// TIA Portal project "PADRAO" (V19)

(* hardware
DEVICE "S7-1200 station_1"  S7-1200 Station
   slot 0: "Rack_0"  S7-1200 Rack  Rack  V1.0
   slot 1: "PLC_1"  CPU 1214C DC/DC/DC  6ES7 214-1AG40-0XB0  V4.4
   slot 2: "DI 8/DQ 8x24VDC_1"  6ES7 223-1BH32-0XB0  V2.0
   slot 3: "CB 1241 (RS485)"  CB 1241 (RS485)  6ES7 241-1CH30-1XB0  V1.0
   slot 3: "DI 8/DQ 8x24VDC_2"  6ES7 223-1BH32-0XB0  V2.0
DEVICE "bb02"  GSD.Device.PN
   slot 0: "Rack"  Rack  V1.0
   slot 0: "bb02"  RT  GMXa-2-Port
      slot 0: "RT"  RT
      slot 1: "bb02"  X1
         slot 1: "Port 1"  Port 1
         slot 2: "Port 2"  Port 2
   slot 1: "Status Device_1"  Status Device
      slot 0: "Status Device"  Status Device
   slot 2: "Device Control_1"  Device Control
      slot 0: "Start/Stop"  Start/Stop
      slot 1: "Reset"  Reset
   slot 3: "Mode_1"  Mode
      slot 0: "Target Mode"  Target Mode
      slot 1: "Operating Mode"  Operating Mode
   slot 4: "Flow Rate_1"  Flow Rate
      slot 0: "Nominal Flow Rate"  Nominal Flow Rate
      slot 1: "Actual Flow Rate"  Actual Flow Rate
   slot 5: "Maximal Flow Rate_1"  Maximal Flow Rate
      slot 0: "Maximal Flow Rate"  Maximal Flow Rate
   slot 9: "Metering Monitor_1"  Metering Monitor
      slot 0: "Metering Monitor"  Metering Monitor
   slot 10: "Error/Warning_1"  Error/Warning
      slot 0: "Error"  Error
      slot 1: "Warning"  Warning
   slot 11: "Strokes/Quantities_1"  Strokes/Quantities
      slot 0: "Reset Stroke Counter"  Reset Stroke Counter
      slot 1: "Reset Quantity Counter"  Reset Quantity Counter
      slot 2: "Stroke Counter"  Stroke Counter
      slot 3: "Quantity Counter"  Quantity Counter
      slot 4: "Litres Per Stroke"  Litres Per Stroke
DEVICE "bb03"  GSD.Device.PN
   slot 0: "Rack"  Rack  V1.0
   slot 0: "bb03"  RT  GMXa-2-Port
      slot 0: "RT"  RT
      slot 1: "bb03"  X1
         slot 1: "Port 1"  Port 1
         slot 2: "Port 2"  Port 2
   slot 1: "Status Device_1"  Status Device
      slot 0: "Status Device"  Status Device
   slot 2: "Device Control_1"  Device Control
      slot 0: "Start/Stop"  Start/Stop
      slot 1: "Reset"  Reset
   slot 3: "Mode_1"  Mode
      slot 0: "Target Mode"  Target Mode
      slot 1: "Operating Mode"  Operating Mode
   slot 4: "Flow Rate_1"  Flow Rate
      slot 0: "Nominal Flow Rate"  Nominal Flow Rate
      slot 1: "Actual Flow Rate"  Actual Flow Rate
   slot 5: "Maximal Flow Rate_1"  Maximal Flow Rate
      slot 0: "Maximal Flow Rate"  Maximal Flow Rate
   slot 9: "Metering Monitor_1"  Metering Monitor
      slot 0: "Metering Monitor"  Metering Monitor
   slot 10: "Error/Warning_1"  Error/Warning
      slot 0: "Error"  Error
      slot 1: "Warning"  Warning
   slot 11: "Strokes/Quantities_1"  Strokes/Quantities
      slot 0: "Reset Stroke Counter"  Reset Stroke Counter
      slot 1: "Reset Quantity Counter"  Reset Quantity Counter
      slot 2: "Stroke Counter"  Stroke Counter
      slot 3: "Quantity Counter"  Quantity Counter
      slot 4: "Litres Per Stroke"  Litres Per Stroke
DEVICE "bb04"  GSD.Device.PN
   slot 0: "Rack"  Rack  V1.0
   slot 0: "bb04"  RT  GMXa-2-Port
      slot 0: "RT"  RT
      slot 1: "bb04"  X1
         slot 1: "Port 1"  Port 1
         slot 2: "Port 2"  Port 2
   slot 1: "Status Device_1"  Status Device
      slot 0: "Status Device"  Status Device
   slot 2: "Device Control_1"  Device Control
      slot 0: "Start/Stop"  Start/Stop
      slot 1: "Reset"  Reset
   slot 3: "Mode_1"  Mode
      slot 0: "Target Mode"  Target Mode
      slot 1: "Operating Mode"  Operating Mode
   slot 4: "Flow Rate_1"  Flow Rate
      slot 0: "Nominal Flow Rate"  Nominal Flow Rate
      slot 1: "Actual Flow Rate"  Actual Flow Rate
   slot 5: "Maximal Flow Rate_1"  Maximal Flow Rate
      slot 0: "Maximal Flow Rate"  Maximal Flow Rate
   slot 9: "Metering Monitor_1"  Metering Monitor
      slot 0: "Metering Monitor"  Metering Monitor
   slot 10: "Error/Warning_1"  Error/Warning
      slot 0: "Error"  Error
      slot 1: "Warning"  Warning
   slot 11: "Strokes/Quantities_1"  Strokes/Quantities
      slot 0: "Reset Stroke Counter"  Reset Stroke Counter
      slot 1: "Reset Quantity Counter"  Reset Quantity Counter
      slot 2: "Stroke Counter"  Stroke Counter
      slot 3: "Quantity Counter"  Quantity Counter
      slot 4: "Litres Per Stroke"  Litres Per Stroke
DEVICE "bb05"  GSD.Device.PN
   slot 0: "Rack"  Rack  V1.0
   slot 0: "bb05"  RT  GMXa-2-Port
      slot 0: "RT"  RT
      slot 1: "bb05"  X1
         slot 1: "Port 1"  Port 1
         slot 2: "Port 2"  Port 2
   slot 1: "Status Device_1"  Status Device
      slot 0: "Status Device"  Status Device
   slot 2: "Device Control_1"  Device Control
      slot 0: "Start/Stop"  Start/Stop
      slot 1: "Reset"  Reset
   slot 3: "Mode_1"  Mode
      slot 0: "Target Mode"  Target Mode
      slot 1: "Operating Mode"  Operating Mode
   slot 4: "Flow Rate_1"  Flow Rate
      slot 0: "Nominal Flow Rate"  Nominal Flow Rate
      slot 1: "Actual Flow Rate"  Actual Flow Rate
   slot 5: "Maximal Flow Rate_1"  Maximal Flow Rate
      slot 0: "Maximal Flow Rate"  Maximal Flow Rate
   slot 9: "Metering Monitor_1"  Metering Monitor
      slot 0: "Metering Monitor"  Metering Monitor
   slot 10: "Error/Warning_1"  Error/Warning
      slot 0: "Error"  Error
      slot 1: "Warning"  Warning
   slot 11: "Strokes/Quantities_1"  Strokes/Quantities
      slot 0: "Reset Stroke Counter"  Reset Stroke Counter
      slot 1: "Reset Quantity Counter"  Reset Quantity Counter
      slot 2: "Stroke Counter"  Stroke Counter
      slot 3: "Quantity Counter"  Quantity Counter
      slot 4: "Litres Per Stroke"  Litres Per Stroke
DEVICE "bb01"  GSD.Device.PN
   slot 0: "Rack"  Rack  V1.0
   slot 0: "bb01"  RT  GMXa-2-Port
      slot 0: "RT"  RT
      slot 1: "bb01"  X1
         slot 1: "Port 1"  Port 1
         slot 2: "Port 2"  Port 2
   slot 1: "Status Device_1"  Status Device
      slot 0: "Status Device"  Status Device
   slot 2: "Device Control_1"  Device Control
      slot 0: "Start/Stop"  Start/Stop
      slot 1: "Reset"  Reset
   slot 3: "Mode_1"  Mode
      slot 0: "Target Mode"  Target Mode
      slot 1: "Operating Mode"  Operating Mode
   slot 4: "Flow Rate_1"  Flow Rate
      slot 0: "Nominal Flow Rate"  Nominal Flow Rate
      slot 1: "Actual Flow Rate"  Actual Flow Rate
   slot 5: "Maximal Flow Rate_1"  Maximal Flow Rate
      slot 0: "Maximal Flow Rate"  Maximal Flow Rate
   slot 9: "Metering Monitor_1"  Metering Monitor
      slot 0: "Metering Monitor"  Metering Monitor
   slot 10: "Error/Warning_1"  Error/Warning
      slot 0: "Error"  Error
      slot 1: "Warning"  Warning
   slot 11: "Strokes/Quantities_1"  Strokes/Quantities
      slot 0: "Reset Stroke Counter"  Reset Stroke Counter
      slot 1: "Reset Quantity Counter"  Reset Quantity Counter
      slot 2: "Stroke Counter"  Stroke Counter
      slot 3: "Quantity Counter"  Quantity Counter
      slot 4: "Litres Per Stroke"  Litres Per Stroke
DEVICE "bb05_1"  GSD.Device.PN
   slot 0: "Rack"  Rack  V1.0
   slot 0: "bb06"  RT  GMXa-2-Port
      slot 0: "RT"  RT
      slot 1: "bb06"  X1
         slot 1: "Port 1"  Port 1
         slot 2: "Port 2"  Port 2
   slot 1: "Status Device_1"  Status Device
      slot 0: "Status Device"  Status Device
   slot 2: "Device Control_1"  Device Control
      slot 0: "Start/Stop"  Start/Stop
      slot 1: "Reset"  Reset
   slot 3: "Mode_1"  Mode
      slot 0: "Target Mode"  Target Mode
      slot 1: "Operating Mode"  Operating Mode
   slot 4: "Flow Rate_1"  Flow Rate
      slot 0: "Nominal Flow Rate"  Nominal Flow Rate
      slot 1: "Actual Flow Rate"  Actual Flow Rate
   slot 5: "Maximal Flow Rate_1"  Maximal Flow Rate
      slot 0: "Maximal Flow Rate"  Maximal Flow Rate
   slot 9: "Metering Monitor_1"  Metering Monitor
      slot 0: "Metering Monitor"  Metering Monitor
   slot 10: "Error/Warning_1"  Error/Warning
      slot 0: "Error"  Error
      slot 1: "Warning"  Warning
   slot 11: "Strokes/Quantities_1"  Strokes/Quantities
      slot 0: "Reset Stroke Counter"  Reset Stroke Counter
      slot 1: "Reset Quantity Counter"  Reset Quantity Counter
      slot 2: "Stroke Counter"  Stroke Counter
      slot 3: "Quantity Counter"  Quantity Counter
      slot 4: "Litres Per Stroke"  Litres Per Stroke
*)

// ===== PLC "PLC_1"  CPU 1214C DC/DC/DC =====

VAR_GLOBAL   // PLC tag table "Default tag table"
   "DI_00" AT %I0.0 : Bool;
   "DI_01" AT %I0.1 : Bool;
   "DI_02" AT %I0.2 : Bool;
   "DI_03" AT %I0.3 : Bool;
   "DI_04" AT %I0.4 : Bool;
   "DI_05" AT %I0.5 : Bool;
   "DI_06" AT %I0.6 : Bool;
   "DI_07" AT %I0.7 : Bool;
   "DI_08" AT %I1.0 : Bool;
   "DI_09" AT %I1.1 : Bool;
   "DI_10" AT %I1.2 : Bool;
   "DI_11" AT %I1.3 : Bool;
   "DI_12" AT %I1.4 : Bool;
   "DI_13" AT %I1.5 : Bool;
   "DO_00" AT %Q0.0 : Bool;
   "DO_01" AT %Q0.1 : Bool;
   "DO_02" AT %Q0.2 : Bool;
   "DO_03" AT %Q0.3 : Bool;
   "DO_04" AT %Q0.4 : Bool;
   "DO_05" AT %Q0.5 : Bool;
   "DO_06" AT %Q0.6 : Bool;
   "DO_07" AT %Q0.7 : Bool;
   "DO_08" AT %Q1.0 : Bool;
   "DO_09" AT %Q1.1 : Bool;
   "System_Byte" AT %MB1 : Byte;
   "FirstScan" AT %M1.0 : Bool;
   "DiagStatusUpdate" AT %M1.1 : Bool;
   "AlwaysTRUE" AT %M1.2 : Bool;
   "AlwaysFALSE" AT %M1.3 : Bool;
   "Clock_Byte" AT %MB0 : Byte;
   "Clock_10Hz" AT %M0.0 : Bool;
   "Clock_5Hz" AT %M0.1 : Bool;
   "Clock_2.5Hz" AT %M0.2 : Bool;
   "Clock_2Hz" AT %M0.3 : Bool;
   "Clock_1.25Hz" AT %M0.4 : Bool;
   "Clock_1Hz" AT %M0.5 : Bool;
   "Clock_0.625Hz" AT %M0.6 : Bool;
   "Clock_0.5Hz" AT %M0.7 : Bool;
   "EmergenciaAcionada" AT %M2.0 : Bool;
   "FaltaFase" AT %M2.1 : Bool;
   "SinalTriturador1" AT %M2.2 : Bool;
   "SinalTriturador2" AT %M2.3 : Bool;
   "SinalMisturador1" AT %M2.4 : Bool;
   "SinalMisturador2" AT %M2.5 : Bool;
   "PulsoMedidor1" AT %M3.3 : Bool;
   "PulsoMedidor2" AT %M3.4 : Bool;
   "PulsoMedidor3" AT %M3.5 : Bool;
   "SistemaHabilitado" AT %M3.6 : Bool;
   "Sirene" AT %M3.7 : Bool;
   "FatorCorrecaoTanque1" AT %MD108 : Real;
   "AI_01" AT %IW64 : Word;
   "AI_02" AT %IW66 : Word;
   "ResetGeral" AT %M4.0 : Bool;
   "VolumePulso1" AT %MD160 : Real;
   "VolumePulso2" AT %MD164 : Real;
   "VolumePulso3" AT %MD172 : Real;
   "NivelBaixoTQ1" AT %M4.1 : Bool;
   "SP_NivelMinimoTanque1" AT %MD184 : Real;
   "StatusFalha" AT %MW192 : Int;
   "FalhaBomba01" AT %M4.5 : Bool;
   "FalhaBomba02" AT %M4.6 : Bool;
   "FalhaBomba03" AT %M4.7 : Bool;
   "FalhaBomba04" AT %M5.0 : Bool;
   "FalhaBomba05" AT %M5.1 : Bool;
   "FatorCorrecaoTanque2" AT %MD112 : Real;
   "SP_NivelMinimoTanque2" AT %MD152 : Real;
   "NivelBaixoTQ2" AT %M7.5 : Bool;
   "LigaValv04" AT %M7.6 : Bool;
   "LigaValv05" AT %M7.7 : Bool;
   "VolumePulso4" AT %MD100 : Real;
   "SP_Dosagem1" AT %MD168 : Real;
   "SP_Dosagem2" AT %MD176 : Real;
   "SP_Dosagem3" AT %MD180 : Real;
   "SP_Dosagem4" AT %MD188 : Real;
   "SP_Dosagem5" AT %MD194 : Real;
   "PulsoMedidor4" AT %M8.2 : Bool;
   "PulsoMedidor5" AT %M8.3 : Bool;
   "FaltaFluxo01" AT %M2.6 : Bool;
   "FaltaFluxo02" AT %M2.7 : Bool;
   "FaltaFluxo03" AT %M3.0 : Bool;
   "FaltaFluxo04" AT %M3.1 : Bool;
   "FaltaFluxo05" AT %M3.2 : Bool;
   "VolumePulso5" AT %MD104 : Real;
   "LigaValv03" AT %M8.0 : Bool;
   "LigaValv06" AT %M8.1 : Bool;
   "RetValvAberta3" AT %M8.5 : Bool;
   "RetValvAberta4" AT %M8.6 : Bool;
   "RetValvAberta5" AT %M8.7 : Bool;
   "RetValvAberta6" AT %M9.0 : Bool;
   "FalhaRetornoValvAberta3" AT %M9.1 : Bool;
   "FalhaRetornoValvAberta4" AT %M9.2 : Bool;
   "FalhaRetornoValvAberta5" AT %M9.3 : Bool;
   "BombaMax1" AT %M4.2 : Bool;
   "BombaMax2" AT %M4.3 : Bool;
   "BombaMax3" AT %M4.4 : Bool;
   "BombaMax4" AT %M5.3 : Bool;
   "BombaMax5" AT %M5.4 : Bool;
   "MedidorEstragado1" AT %M5.5 : Bool;
   "MedidorEstragado2" AT %M5.6 : Bool;
   "MedidorEstragado3" AT %M5.7 : Bool;
   "MedidorEstragado4" AT %M6.0 : Bool;
   "MedidorEstragado5" AT %M6.1 : Bool;
   "IniciaCalibracao1" AT %M6.3 : Bool;
   "IniciaCalibracao2" AT %M6.4 : Bool;
   "IniciaCalibracao3" AT %M6.5 : Bool;
   "IniciaCalibracao4" AT %M6.6 : Bool;
   "IniciaCalibracao5" AT %M6.7 : Bool;
   "BombaMax6" AT %M7.1 : Bool;
   "FalhaBomba06" AT %M5.2 : Bool;
   "FalhaRetornoValvAberta6" AT %M9.4 : Bool;
   "FaltaFluxo06" AT %M6.2 : Bool;
   "VolumePulso6" AT %MD116 : Real;
   "IniciaCalibracao6" AT %M7.0 : Bool;
   "MedidorEstragado6" AT %M7.2 : Bool;
   "PulsoMedidor6" AT %M8.4 : Bool;
   "SP_Dosagem6" AT %MD198 : Real;
   "SP_NivelMuitoBaixoTanque1" AT %MD120 : Real;
   "SP_NivelMuitoBaixoTanque2" AT %MD124 : Real;
   "NivelMuitoBaixoTQ1" AT %M7.3 : Bool;
   "NivelMuitoBaixoTQ2" AT %M7.4 : Bool;
   "OffSetTQ1" AT %MD128 : Real;
   "OffSetTQ2" AT %MD132 : Real;
   "CircunferenciaTQ1" AT %MD136 : Real;
   "CircunferenciaTQ2" AT %MD140 : Real;
   "StatusBombaEspelho" AT %MD144 : DInt;
   "DataEspelho" AT %MD148 : DInt;
   "HoraEspelho" AT %MD156 : DInt;
   "DI_14" AT %I8.0 : Bool;
   "DI_15" AT %I8.1 : Bool;
   "DI_16" AT %I8.2 : Bool;
   "DI_17" AT %I8.3 : Bool;
   "DI_18" AT %I8.4 : Bool;
   "DI_19" AT %I8.5 : Bool;
   "DI_20" AT %I8.6 : Bool;
   "DI_21" AT %I8.7 : Bool;
   "SP_DelayFinal1" AT %MD202 : Time;
   "SP_DelayFinal2" AT %MD206 : Time;
   "SP_DelayFinal3" AT %MD210 : Time;
   "SP_DelayFinal4" AT %MD214 : Time;
   "SP_DelayFinal5" AT %MD218 : Time;
   "SP_DelayFinal6" AT %MD222 : Time;
   "FalhaRetBomba1" AT %M9.5 : Bool;
   "FalhaRetBomba2" AT %M9.6 : Bool;
   "FalhaRetBomba3" AT %M9.7 : Bool;
   "FalhaRetBomba4" AT %M10.0 : Bool;
   "FalhaRetBomba5" AT %M10.1 : Bool;
   "FalhaRetBomba6" AT %M10.2 : Bool;
   "QuedaEnergia" AT %M10.3 : Bool;
   "Frequencia1" AT %MD246 : Real;
   "SP_DelayIniciaPID" AT %MD242 : Time;
   "Frequencia2" AT %MD250 : Real;
   "Frequencia3" AT %MD254 : Real;
   "Frequencia4" AT %MD258 : Real;
   "Frequencia5" AT %MD262 : Real;
   "Frequencia6" AT %MD300 : Real;
   "SP_DelayColaFreq" AT %MD12 : Time;
END_VAR

// folder: Common

TYPE "typeDiagnostics"
TITLE = typeDiagnostics
// Provides a structure for detailed diagnostics
   STRUCT
      status : Word;   // Status of the block or error identification when error occurred
      subfunctionStatus : DWord;   // Status or return value of called FBs, FCs and system blocks
      stateNumber : DInt;   // State in the state machine of the block where the error occurred
   END_STRUCT;
END_TYPE

// folder: LMQTT

TYPE "LMQTT_typeConnParam"
TITLE = LMQTT_typeConnParams
// Specifies connection parameters for the mqtt connection
   STRUCT
      hwId : Hw_Any;   // Hardware identifier of the interface. 0: interface is selected automatically
      connId : Conn_Ouc := 1;   // Unique connection identifier (1..4095)
      broker : String;   // Hostname or IP address of broker
      port : UInt := 1883;   // Port on the broker
      tls : Struct   // Parameters for TLS encryption
         enableTls : Bool;   // TRUE: Enables TLS, FALSE: disable TLS
         validateServerIdentity : Bool;   // TRUE: Validate server certificate, FALSE: No validation of server certificate
         brokerCert : UDInt;   // ID of the broker's certificate in TIA Portal
         clientCert : UDInt;   // ID of the client's certificate in TIA Portal
      END_STRUCT;
      keepAlive : UInt;   // Keepalive mechanism for MQTT in seconds. 0: disabled.
   END_STRUCT;
END_TYPE

// folder: DB

DATA_BLOCK "RelatorioUnificado"   // DB1
{ S7_Optimized_Access := 'TRUE' }
VERSION : 0.1
   VAR RETAIN
      Diario : Array[1..20] of Real;
      Totalizador : Array[1..20] of Real;
      DosagemAtual : Array[1..20] of Real;
   END_VAR
BEGIN
END_DATA_BLOCK

DATA_BLOCK "InputClp_DB"   // DB2
{ S7_Optimized_Access := 'TRUE' }
VERSION : 0.1
// stored: InstanceOfName InputClp
"InputClp"
BEGIN
END_DATA_BLOCK

DATA_BLOCK "NivelTanque1"   // DB3
{ S7_Optimized_Access := 'TRUE' }
VERSION : 0.1
// stored: InstanceOfName NivelTanque
"NivelTanque"
BEGIN
END_DATA_BLOCK

DATA_BLOCK "InputClp_DB2"   // DB4
{ S7_Optimized_Access := 'TRUE' }
VERSION : 0.1
// stored: InstanceOfName InputClp
"InputClp"
BEGIN
END_DATA_BLOCK

DATA_BLOCK "OutputClp_DB"   // DB5
{ S7_Optimized_Access := 'TRUE' }
VERSION : 0.1
// stored: InstanceOfName OutputClp
"OutputClp"
BEGIN
END_DATA_BLOCK

DATA_BLOCK "NivelTanque2"   // DB6
{ S7_Optimized_Access := 'TRUE' }
VERSION : 0.1
// stored: InstanceOfName NivelTanque
"NivelTanque"
BEGIN
END_DATA_BLOCK

DATA_BLOCK "DosagemContinua_DB1"   // DB7
{ S7_Optimized_Access := 'TRUE' }
VERSION : 0.1
// stored: InstanceOfName DosagemContinua
"DosagemContinua"
BEGIN
END_DATA_BLOCK

DATA_BLOCK "RegistradorMedidor_DB1"   // DB8
{ S7_Optimized_Access := 'TRUE' }
VERSION : 0.1
// stored: InstanceOfName RegistradorMedidor
"RegistradorMedidor"
BEGIN
END_DATA_BLOCK

DATA_BLOCK "DosagemContinua_DB2"   // DB9
{ S7_Optimized_Access := 'TRUE' }
VERSION : 0.1
// stored: InstanceOfName DosagemContinua
"DosagemContinua"
BEGIN
END_DATA_BLOCK

DATA_BLOCK "RegistradorMedidor_DB2"   // DB10
{ S7_Optimized_Access := 'TRUE' }
VERSION : 0.1
// stored: InstanceOfName RegistradorMedidor
"RegistradorMedidor"
BEGIN
END_DATA_BLOCK

DATA_BLOCK "DosagemContinua_DB3"   // DB11
{ S7_Optimized_Access := 'TRUE' }
VERSION : 0.1
// stored: InstanceOfName DosagemContinua
"DosagemContinua"
BEGIN
END_DATA_BLOCK

DATA_BLOCK "RegistradorMedidor_DB3"   // DB12
{ S7_Optimized_Access := 'TRUE' }
VERSION : 0.1
// stored: InstanceOfName RegistradorMedidor
"RegistradorMedidor"
BEGIN
END_DATA_BLOCK

DATA_BLOCK "DosagemContinua_DB4"   // DB13
{ S7_Optimized_Access := 'TRUE' }
VERSION : 0.1
// stored: InstanceOfName DosagemContinua
"DosagemContinua"
BEGIN
END_DATA_BLOCK

DATA_BLOCK "RelatorioSAPI"   // DB14
{ S7_Optimized_Access := 'TRUE' }
VERSION : 0.1
   VAR RETAIN
      Hora : Array[1..200] of Real;
      TotalTempoBomba : Array[1..20] of DInt;
      TotalTempoSinal : Array[1..20] of DInt;
      TotalAcionamentosSinal : Array[1..20] of DInt;
      TotalAcionamentosBBA : Array[1..20] of DInt;
      auxPulsoClock : Array[1..40] of Bool;
      auxNegaSinal : Array[1..20] of Bool;
      auxNegaBomba : Array[1..20] of Bool;
      StatusINT : Int := -1;
      StatusReal : Real := -1.0;
   END_VAR
   VAR
      GravaFTP : Bool;
      EnviaFTP : Bool;
      TesteGrava : Bool;
      TesteEnvia : Bool;
      TesteSet : Bool;
   END_VAR
BEGIN
   Hora[1] := -1.0;
   Hora[2] := -1.0;
   Hora[3] := -1.0;
   Hora[4] := -1.0;
   Hora[5] := -1.0;
   Hora[6] := -1.0;
   Hora[7] := -1.0;
   Hora[8] := -1.0;
   Hora[9] := -1.0;
   Hora[10] := -1.0;
   Hora[11] := -1.0;
   Hora[12] := -1.0;
   Hora[13] := -1.0;
   Hora[14] := -1.0;
   Hora[15] := -1.0;
   Hora[16] := -1.0;
   Hora[17] := -1.0;
   Hora[18] := -1.0;
   Hora[19] := -1.0;
   Hora[20] := -1.0;
   Hora[21] := -1.0;
   Hora[22] := -1.0;
   Hora[23] := -1.0;
   Hora[24] := -1.0;
   Hora[25] := -1.0;
   Hora[26] := -1.0;
   Hora[27] := -1.0;
   Hora[28] := -1.0;
   Hora[29] := -1.0;
   Hora[30] := -1.0;
   Hora[31] := -1.0;
   Hora[32] := -1.0;
   Hora[33] := -1.0;
   Hora[34] := -1.0;
   Hora[35] := -1.0;
   Hora[36] := -1.0;
   Hora[37] := -1.0;
   Hora[38] := -1.0;
   Hora[39] := -1.0;
   Hora[40] := -1.0;
   Hora[41] := -1.0;
   Hora[42] := -1.0;
   Hora[43] := -1.0;
   Hora[44] := -1.0;
   Hora[45] := -1.0;
   Hora[46] := -1.0;
   Hora[47] := -1.0;
   Hora[48] := -1.0;
   Hora[49] := -1.0;
   Hora[50] := -1.0;
   Hora[51] := -1.0;
   Hora[52] := -1.0;
   Hora[53] := -1.0;
   Hora[54] := -1.0;
   Hora[55] := -1.0;
   Hora[56] := -1.0;
   Hora[57] := -1.0;
   Hora[58] := -1.0;
   Hora[59] := -1.0;
   Hora[60] := -1.0;
   Hora[61] := -1.0;
   Hora[62] := -1.0;
   Hora[63] := -1.0;
   Hora[64] := -1.0;
   Hora[65] := -1.0;
   Hora[66] := -1.0;
   Hora[67] := -1.0;
   Hora[68] := -1.0;
   Hora[69] := -1.0;
   Hora[70] := -1.0;
   Hora[71] := -1.0;
   Hora[72] := -1.0;
   Hora[73] := -1.0;
   Hora[74] := -1.0;
   Hora[75] := -1.0;
   Hora[76] := -1.0;
   Hora[77] := -1.0;
   Hora[78] := -1.0;
   Hora[79] := -1.0;
   Hora[80] := -1.0;
   Hora[81] := -1.0;
   Hora[82] := -1.0;
   Hora[83] := -1.0;
   Hora[84] := -1.0;
   Hora[85] := -1.0;
   Hora[86] := -1.0;
   Hora[87] := -1.0;
   Hora[88] := -1.0;
   Hora[89] := -1.0;
   Hora[90] := -1.0;
   Hora[91] := -1.0;
   Hora[92] := -1.0;
   Hora[93] := -1.0;
   Hora[94] := -1.0;
   Hora[95] := -1.0;
   Hora[96] := -1.0;
   Hora[97] := -1.0;
   Hora[98] := -1.0;
   Hora[99] := -1.0;
   Hora[100] := -1.0;
   Hora[101] := -1.0;
   Hora[102] := -1.0;
   Hora[103] := -1.0;
   Hora[104] := -1.0;
   Hora[105] := -1.0;
   Hora[106] := -1.0;
   Hora[107] := -1.0;
   Hora[108] := -1.0;
   Hora[109] := -1.0;
   Hora[110] := -1.0;
   Hora[111] := -1.0;
   Hora[112] := -1.0;
   Hora[113] := -1.0;
   Hora[114] := -1.0;
   Hora[115] := -1.0;
   Hora[116] := -1.0;
   Hora[117] := -1.0;
   Hora[118] := -1.0;
   Hora[119] := -1.0;
   Hora[120] := -1.0;
   Hora[121] := -1.0;
   Hora[122] := -1.0;
   Hora[123] := -1.0;
   Hora[124] := -1.0;
   Hora[125] := -1.0;
   Hora[126] := -1.0;
   Hora[127] := -1.0;
   Hora[128] := -1.0;
   Hora[129] := -1.0;
   Hora[130] := -1.0;
   Hora[131] := -1.0;
   Hora[132] := -1.0;
   Hora[133] := -1.0;
   Hora[134] := -1.0;
   Hora[135] := -1.0;
   Hora[136] := -1.0;
   Hora[137] := -1.0;
   Hora[138] := -1.0;
   Hora[139] := -1.0;
   Hora[140] := -1.0;
   Hora[141] := -1.0;
   Hora[142] := -1.0;
   Hora[143] := -1.0;
   Hora[144] := -1.0;
   Hora[145] := -1.0;
   Hora[146] := -1.0;
   Hora[147] := -1.0;
   Hora[148] := -1.0;
   Hora[149] := -1.0;
   Hora[150] := -1.0;
   Hora[151] := -1.0;
   Hora[152] := -1.0;
   Hora[153] := -1.0;
   Hora[154] := -1.0;
   Hora[155] := -1.0;
   Hora[156] := -1.0;
   Hora[157] := -1.0;
   Hora[158] := -1.0;
   Hora[159] := -1.0;
   Hora[160] := -1.0;
   Hora[161] := -1.0;
   Hora[162] := -1.0;
   Hora[163] := -1.0;
   Hora[164] := -1.0;
   Hora[165] := -1.0;
   Hora[166] := -1.0;
   Hora[167] := -1.0;
   Hora[168] := -1.0;
   Hora[169] := -1.0;
   Hora[170] := -1.0;
   Hora[171] := -1.0;
   Hora[172] := -1.0;
   Hora[173] := -1.0;
   Hora[174] := -1.0;
   Hora[175] := -1.0;
   Hora[176] := -1.0;
   Hora[177] := -1.0;
   Hora[178] := -1.0;
   Hora[179] := -1.0;
   Hora[180] := -1.0;
   Hora[181] := -1.0;
   Hora[182] := -1.0;
   Hora[183] := -1.0;
   Hora[184] := -1.0;
   Hora[185] := -1.0;
   Hora[186] := -1.0;
   Hora[187] := -1.0;
   Hora[188] := -1.0;
   Hora[189] := -1.0;
   Hora[190] := -1.0;
   Hora[191] := -1.0;
   Hora[192] := -1.0;
   Hora[193] := -1.0;
   Hora[194] := -1.0;
   Hora[195] := -1.0;
   Hora[196] := -1.0;
   Hora[197] := -1.0;
   Hora[198] := -1.0;
   Hora[199] := -1.0;
   Hora[200] := -1.0;
END_DATA_BLOCK

DATA_BLOCK "RegistradorMedidor_DB4"   // DB15
{ S7_Optimized_Access := 'TRUE' }
VERSION : 0.1
// stored: InstanceOfName RegistradorMedidor
"RegistradorMedidor"
BEGIN
END_DATA_BLOCK

DATA_BLOCK "InterfaceProfi1"   // DB16
{ S7_Optimized_Access := 'TRUE' }
AUTHOR : kellerc
FAMILY : GammaX
NAME : Basic
VERSION : 1.0
// stored: InstanceOfName FBGammaX_1200
"FBGammaX_1200"
BEGIN
END_DATA_BLOCK

DATA_BLOCK "DosagemContinua_DB5"   // DB17
{ S7_Optimized_Access := 'TRUE' }
VERSION : 0.1
// stored: InstanceOfName DosagemContinua
"DosagemContinua"
BEGIN
END_DATA_BLOCK

DATA_BLOCK "InterfaceProfi2"   // DB18
{ S7_Optimized_Access := 'TRUE' }
AUTHOR : kellerc
FAMILY : GammaX
NAME : Basic
VERSION : 1.0
// stored: InstanceOfName FBGammaX_1200
"FBGammaX_1200"
BEGIN
END_DATA_BLOCK

DATA_BLOCK "InterfaceProfi3"   // DB19
{ S7_Optimized_Access := 'TRUE' }
AUTHOR : kellerc
FAMILY : GammaX
NAME : Basic
VERSION : 1.0
// stored: InstanceOfName FBGammaX_1200
"FBGammaX_1200"
BEGIN
END_DATA_BLOCK

DATA_BLOCK "InterfaceProfi4"   // DB20
{ S7_Optimized_Access := 'TRUE' }
AUTHOR : kellerc
FAMILY : GammaX
NAME : Basic
VERSION : 1.0
// stored: InstanceOfName FBGammaX_1200
"FBGammaX_1200"
BEGIN
END_DATA_BLOCK

DATA_BLOCK "InterfaceProfi5"   // DB21
{ S7_Optimized_Access := 'TRUE' }
AUTHOR : kellerc
FAMILY : GammaX
NAME : Basic
VERSION : 1.0
// stored: InstanceOfName FBGammaX_1200
"FBGammaX_1200"
BEGIN
END_DATA_BLOCK

DATA_BLOCK "RegistradorMedidor_DB5"   // DB22
{ S7_Optimized_Access := 'TRUE' }
VERSION : 0.1
// stored: InstanceOfName RegistradorMedidor
"RegistradorMedidor"
BEGIN
END_DATA_BLOCK

DATA_BLOCK "DosagemContinua_DB6"   // DB23
{ S7_Optimized_Access := 'TRUE' }
VERSION : 0.1
// stored: InstanceOfName DosagemContinua
"DosagemContinua"
BEGIN
END_DATA_BLOCK

DATA_BLOCK "RegistradorMedidor_DB6"   // DB24
{ S7_Optimized_Access := 'TRUE' }
VERSION : 0.1
// stored: InstanceOfName RegistradorMedidor
"RegistradorMedidor"
BEGIN
END_DATA_BLOCK

DATA_BLOCK "InterfaceProfi6"   // DB31
{ S7_Optimized_Access := 'TRUE' }
AUTHOR : kellerc
FAMILY : GammaX
NAME : Basic
VERSION : 1.0
// stored: InstanceOfName FBGammaX_1200
"FBGammaX_1200"
BEGIN
END_DATA_BLOCK

DATA_BLOCK "DataTime"   // DB48
{ S7_Optimized_Access := 'TRUE' }
VERSION : 0.1
   VAR RETAIN
      DataHora : DTL;
      IHM : Array[0..6] of Word;
   END_VAR
BEGIN
END_DATA_BLOCK

DATA_BLOCK "SetDbSapi_DB"   // DB87
{ S7_Optimized_Access := 'TRUE' }
VERSION : 0.1
// stored: InstanceOfName SetDbSapi
"SetDbSapi"
BEGIN
END_DATA_BLOCK

// folder: System blocks/Program resources

DATA_BLOCK "TON_FalhaRetornoValv3"   // DB25
{ S7_Optimized_Access := 'TRUE' }
AUTHOR : Simatic
FAMILY : IEC
NAME : IEC_TMR
VERSION : 1.0
// stored: InstanceOfName IEC_TIMER
"IEC_TIMER"
BEGIN
END_DATA_BLOCK

DATA_BLOCK "TON_FalhaRetornoValv4"   // DB26
{ S7_Optimized_Access := 'TRUE' }
AUTHOR : Simatic
FAMILY : IEC
NAME : IEC_TMR
VERSION : 1.0
// stored: InstanceOfName IEC_TIMER
"IEC_TIMER"
BEGIN
END_DATA_BLOCK

DATA_BLOCK "TON_FalhaRetornoValv5"   // DB27
{ S7_Optimized_Access := 'TRUE' }
AUTHOR : Simatic
FAMILY : IEC
NAME : IEC_TMR
VERSION : 1.0
// stored: InstanceOfName IEC_TIMER
"IEC_TIMER"
BEGIN
END_DATA_BLOCK

DATA_BLOCK "TON_FalhaRetornoValv6"   // DB28
{ S7_Optimized_Access := 'TRUE' }
AUTHOR : Simatic
FAMILY : IEC
NAME : IEC_TMR
VERSION : 1.0
// stored: InstanceOfName IEC_TIMER
"IEC_TIMER"
BEGIN
END_DATA_BLOCK

DATA_BLOCK "TON_DelayIniciaPID1"   // DB29
{ S7_Optimized_Access := 'TRUE' }
AUTHOR : Simatic
FAMILY : IEC
NAME : IEC_TMR
VERSION : 1.0
// stored: InstanceOfName IEC_TIMER
"IEC_TIMER"
BEGIN
END_DATA_BLOCK

DATA_BLOCK "TON_DelayIniciaPID2"   // DB30
{ S7_Optimized_Access := 'TRUE' }
AUTHOR : Simatic
FAMILY : IEC
NAME : IEC_TMR
VERSION : 1.0
// stored: InstanceOfName IEC_TIMER
"IEC_TIMER"
BEGIN
END_DATA_BLOCK

DATA_BLOCK "TON_DelayIniciaPID3"   // DB32
{ S7_Optimized_Access := 'TRUE' }
AUTHOR : Simatic
FAMILY : IEC
NAME : IEC_TMR
VERSION : 1.0
// stored: InstanceOfName IEC_TIMER
"IEC_TIMER"
BEGIN
END_DATA_BLOCK

DATA_BLOCK "TON_DelayIniciaPID4"   // DB33
{ S7_Optimized_Access := 'TRUE' }
AUTHOR : Simatic
FAMILY : IEC
NAME : IEC_TMR
VERSION : 1.0
// stored: InstanceOfName IEC_TIMER
"IEC_TIMER"
BEGIN
END_DATA_BLOCK

DATA_BLOCK "TON_DelayIniciaPID5"   // DB34
{ S7_Optimized_Access := 'TRUE' }
AUTHOR : Simatic
FAMILY : IEC
NAME : IEC_TMR
VERSION : 1.0
// stored: InstanceOfName IEC_TIMER
"IEC_TIMER"
BEGIN
END_DATA_BLOCK

DATA_BLOCK "TON_DelayIniciaPID6"   // DB35
{ S7_Optimized_Access := 'TRUE' }
AUTHOR : Simatic
FAMILY : IEC
NAME : IEC_TMR
VERSION : 1.0
// stored: InstanceOfName IEC_TIMER
"IEC_TIMER"
BEGIN
END_DATA_BLOCK

DATA_BLOCK "TON_ResetQuedaEnergia"   // DB42
{ S7_Optimized_Access := 'TRUE' }
AUTHOR : Simatic
FAMILY : IEC
NAME : IEC_TMR
VERSION : 1.0
// stored: InstanceOfName IEC_TIMER
"IEC_TIMER"
BEGIN
END_DATA_BLOCK

DATA_BLOCK "TOF_ResetGeral"   // DB43
{ S7_Optimized_Access := 'TRUE' }
AUTHOR : Simatic
FAMILY : IEC
NAME : IEC_TMR
VERSION : 1.0
// stored: InstanceOfName IEC_TIMER
"IEC_TIMER"
BEGIN
END_DATA_BLOCK

DATA_BLOCK "ModbusTimer1"   // DB46
{ S7_Optimized_Access := 'TRUE' }
AUTHOR : Simatic
FAMILY : IEC
NAME : IEC_TMR
VERSION : 1.0
// stored: InstanceOfName IEC_TIMER
"IEC_TIMER"
BEGIN
END_DATA_BLOCK

DATA_BLOCK "ContadorFalha1"   // DB47
{ S7_Optimized_Access := 'TRUE' }
AUTHOR : Simatic
FAMILY : IEC
NAME : CNTR
VERSION : 1.0
// stored: InstanceOfName IEC_COUNTER
"IEC_COUNTER"
BEGIN
END_DATA_BLOCK

DATA_BLOCK "TON_FaltaFluxo1"   // DB49
{ S7_Optimized_Access := 'TRUE' }
AUTHOR : Simatic
FAMILY : IEC
NAME : IEC_TMR
VERSION : 1.0
// stored: InstanceOfName IEC_TIMER
"IEC_TIMER"
BEGIN
END_DATA_BLOCK

DATA_BLOCK "ContadorFalha2"   // DB50
{ S7_Optimized_Access := 'TRUE' }
AUTHOR : Simatic
FAMILY : IEC
NAME : CNTR
VERSION : 1.0
// stored: InstanceOfName IEC_COUNTER
"IEC_COUNTER"
BEGIN
END_DATA_BLOCK

DATA_BLOCK "T2_FalhaComunicacaoNexxus"   // DB51
{ S7_Optimized_Access := 'TRUE' }
AUTHOR : Simatic
FAMILY : IEC
NAME : IEC_TMR
VERSION : 1.0
// stored: InstanceOfName IEC_TIMER
"IEC_TIMER"
BEGIN
END_DATA_BLOCK

DATA_BLOCK "TON_FaltaFluxo2"   // DB53
{ S7_Optimized_Access := 'TRUE' }
AUTHOR : Simatic
FAMILY : IEC
NAME : IEC_TMR
VERSION : 1.0
// stored: InstanceOfName IEC_TIMER
"IEC_TIMER"
BEGIN
END_DATA_BLOCK

DATA_BLOCK "TON_FaltaFluxo3"   // DB54
{ S7_Optimized_Access := 'TRUE' }
AUTHOR : Simatic
FAMILY : IEC
NAME : IEC_TMR
VERSION : 1.0
// stored: InstanceOfName IEC_TIMER
"IEC_TIMER"
BEGIN
END_DATA_BLOCK

DATA_BLOCK "TON_FaltaFluxo6"   // DB63
{ S7_Optimized_Access := 'TRUE' }
AUTHOR : Simatic
FAMILY : IEC
NAME : IEC_TMR
VERSION : 1.0
// stored: InstanceOfName IEC_TIMER
"IEC_TIMER"
BEGIN
END_DATA_BLOCK

DATA_BLOCK "T1_FalhaComunicacaoNexxu1"   // DB64
{ S7_Optimized_Access := 'TRUE' }
AUTHOR : Simatic
FAMILY : IEC
NAME : IEC_TMR
VERSION : 1.0
// stored: InstanceOfName IEC_TIMER
"IEC_TIMER"
BEGIN
END_DATA_BLOCK

DATA_BLOCK "TON_FaltaFluxo4"   // DB65
{ S7_Optimized_Access := 'TRUE' }
AUTHOR : Simatic
FAMILY : IEC
NAME : IEC_TMR
VERSION : 1.0
// stored: InstanceOfName IEC_TIMER
"IEC_TIMER"
BEGIN
END_DATA_BLOCK

DATA_BLOCK "TON_FaltaFluxo5"   // DB66
{ S7_Optimized_Access := 'TRUE' }
AUTHOR : Simatic
FAMILY : IEC
NAME : IEC_TMR
VERSION : 1.0
// stored: InstanceOfName IEC_TIMER
"IEC_TIMER"
BEGIN
END_DATA_BLOCK

DATA_BLOCK "TON_FalhaRetorno3"   // DB76
{ S7_Optimized_Access := 'TRUE' }
AUTHOR : Simatic
FAMILY : IEC
NAME : IEC_TMR
VERSION : 1.0
// stored: InstanceOfName IEC_TIMER
"IEC_TIMER"
BEGIN
END_DATA_BLOCK

DATA_BLOCK "TON_FalhaRetorno2"   // DB77
{ S7_Optimized_Access := 'TRUE' }
AUTHOR : Simatic
FAMILY : IEC
NAME : IEC_TMR
VERSION : 1.0
// stored: InstanceOfName IEC_TIMER
"IEC_TIMER"
BEGIN
END_DATA_BLOCK

DATA_BLOCK "TON_FalhaRetorno1"   // DB78
{ S7_Optimized_Access := 'TRUE' }
AUTHOR : Simatic
FAMILY : IEC
NAME : IEC_TMR
VERSION : 1.0
// stored: InstanceOfName IEC_TIMER
"IEC_TIMER"
BEGIN
END_DATA_BLOCK

DATA_BLOCK "TON_FalhaRetorno5"   // DB79
{ S7_Optimized_Access := 'TRUE' }
AUTHOR : Simatic
FAMILY : IEC
NAME : IEC_TMR
VERSION : 1.0
// stored: InstanceOfName IEC_TIMER
"IEC_TIMER"
BEGIN
END_DATA_BLOCK

DATA_BLOCK "TON_FalhaRetorno6"   // DB80
{ S7_Optimized_Access := 'TRUE' }
AUTHOR : Simatic
FAMILY : IEC
NAME : IEC_TMR
VERSION : 1.0
// stored: InstanceOfName IEC_TIMER
"IEC_TIMER"
BEGIN
END_DATA_BLOCK

DATA_BLOCK "TON_FalhaRetorno4"   // DB81
{ S7_Optimized_Access := 'TRUE' }
AUTHOR : Simatic
FAMILY : IEC
NAME : IEC_TMR
VERSION : 1.0
// stored: InstanceOfName IEC_TIMER
"IEC_TIMER"
BEGIN
END_DATA_BLOCK

// folder: (top level)

ORGANIZATION_BLOCK "07-PID"   // OB30, LAD, CyclicInterrupt
{ S7_Optimized_Access := 'TRUE' }
VERSION : 0.1
   VAR_INPUT
      Initial_Call : Bool;   // Initial call of this OB
      Event_Count : Int;   // Events discarded
   END_VAR
BEGIN

REGION Network 1: PID 1
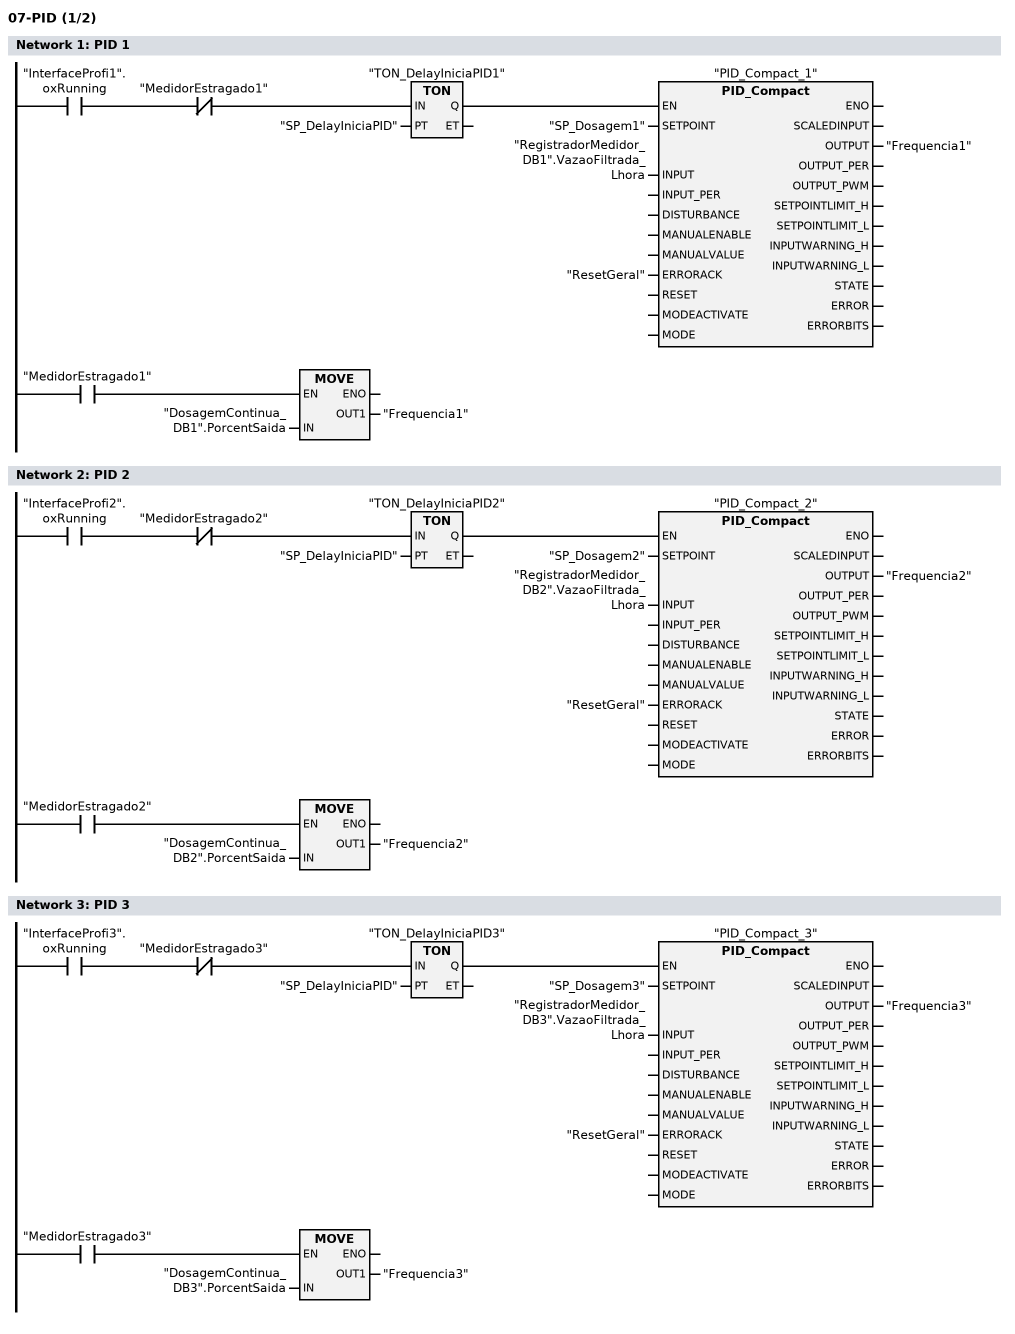
   "TON_DelayIniciaPID1".TON(IN := "InterfaceProfi1".oxRunning AND NOT "MedidorEstragado1",
                           PT := "SP_DelayIniciaPID");
   IF "TON_DelayIniciaPID1".Q THEN
       "PID_Compact_1"(Setpoint := "SP_Dosagem1",   // PID_Compact
                       Input := "RegistradorMedidor_DB1".VazaoFiltrada_Lhora,
                       ErrorAck := "ResetGeral",
                       Output => "Frequencia1");
   END_IF;
   IF "MedidorEstragado1" THEN "Frequencia1" := "DosagemContinua_DB1".PorcentSaida; END_IF;
END_REGION

REGION Network 2: PID 2
   "TON_DelayIniciaPID2".TON(IN := "InterfaceProfi2".oxRunning AND NOT "MedidorEstragado2",
                           PT := "SP_DelayIniciaPID");
   IF "TON_DelayIniciaPID2".Q THEN
       "PID_Compact_2"(Setpoint := "SP_Dosagem2",   // PID_Compact
                       Input := "RegistradorMedidor_DB2".VazaoFiltrada_Lhora,
                       ErrorAck := "ResetGeral",
                       Output => "Frequencia2");
   END_IF;
   IF "MedidorEstragado2" THEN "Frequencia2" := "DosagemContinua_DB2".PorcentSaida; END_IF;
END_REGION

REGION Network 3: PID 3
   "TON_DelayIniciaPID3".TON(IN := "InterfaceProfi3".oxRunning AND NOT "MedidorEstragado3",
                           PT := "SP_DelayIniciaPID");
   IF "TON_DelayIniciaPID3".Q THEN
       "PID_Compact_3"(Setpoint := "SP_Dosagem3",   // PID_Compact
                       Input := "RegistradorMedidor_DB3".VazaoFiltrada_Lhora,
                       ErrorAck := "ResetGeral",
                       Output => "Frequencia3");
   END_IF;
   IF "MedidorEstragado3" THEN "Frequencia3" := "DosagemContinua_DB3".PorcentSaida; END_IF;
END_REGION

REGION Network 4: PID 4
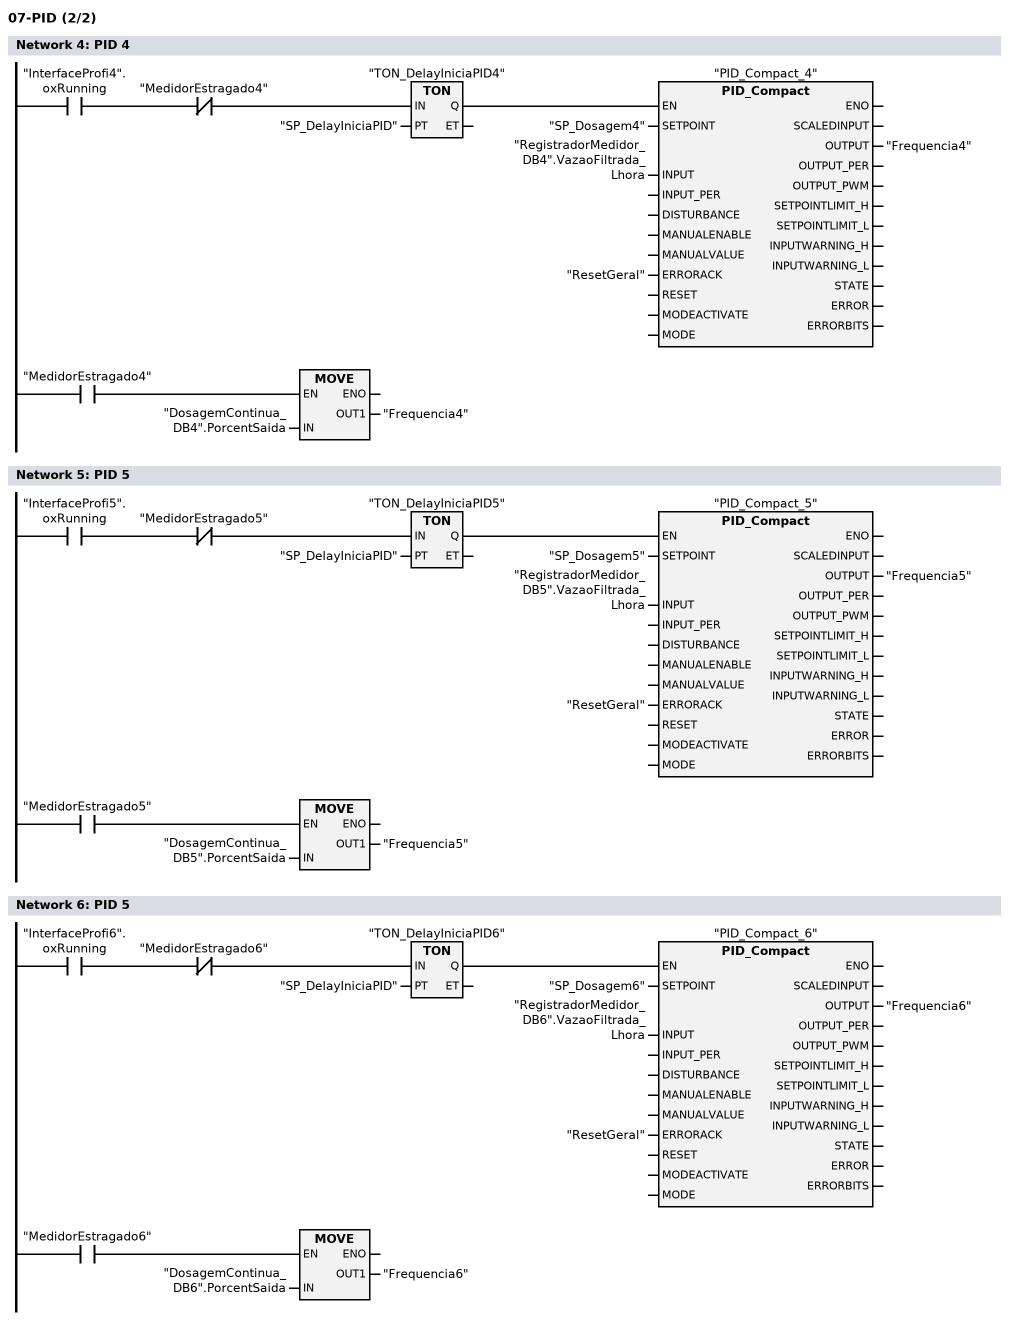
   "TON_DelayIniciaPID4".TON(IN := "InterfaceProfi4".oxRunning AND NOT "MedidorEstragado4",
                           PT := "SP_DelayIniciaPID");
   IF "TON_DelayIniciaPID4".Q THEN
       "PID_Compact_4"(Setpoint := "SP_Dosagem4",   // PID_Compact
                       Input := "RegistradorMedidor_DB4".VazaoFiltrada_Lhora,
                       ErrorAck := "ResetGeral",
                       Output => "Frequencia4");
   END_IF;
   IF "MedidorEstragado4" THEN "Frequencia4" := "DosagemContinua_DB4".PorcentSaida; END_IF;
END_REGION

REGION Network 5: PID 5
   "TON_DelayIniciaPID5".TON(IN := "InterfaceProfi5".oxRunning AND NOT "MedidorEstragado5",
                           PT := "SP_DelayIniciaPID");
   IF "TON_DelayIniciaPID5".Q THEN
       "PID_Compact_5"(Setpoint := "SP_Dosagem5",   // PID_Compact
                       Input := "RegistradorMedidor_DB5".VazaoFiltrada_Lhora,
                       ErrorAck := "ResetGeral",
                       Output => "Frequencia5");
   END_IF;
   IF "MedidorEstragado5" THEN "Frequencia5" := "DosagemContinua_DB5".PorcentSaida; END_IF;
END_REGION

REGION Network 6: PID 5
   "TON_DelayIniciaPID6".TON(IN := "InterfaceProfi6".oxRunning AND NOT "MedidorEstragado6",
                           PT := "SP_DelayIniciaPID");
   IF "TON_DelayIniciaPID6".Q THEN
       "PID_Compact_6"(Setpoint := "SP_Dosagem6",   // PID_Compact
                       Input := "RegistradorMedidor_DB6".VazaoFiltrada_Lhora,
                       ErrorAck := "ResetGeral",
                       Output => "Frequencia6");
   END_IF;
   IF "MedidorEstragado6" THEN "Frequencia6" := "DosagemContinua_DB6".PorcentSaida; END_IF;
END_REGION
END_ORGANIZATION_BLOCK

ORGANIZATION_BLOCK "01-EspelhoInOut"   // OB123, LAD, ProgramCycle
TITLE = "Main Program Sweep (Cycle)"
{ S7_Optimized_Access := 'TRUE' }
VERSION : 0.1
// Espelho das entradas e saidas do CLP
   VAR_INPUT
      Initial_Call : Bool;   // Initial call of this OB
      Remanence : Bool;   // =True, if remanent data are available
   END_VAR
   VAR_TEMP   // added for the SCL form of the ladder/FBD networks
      _w1 : Bool;
   END_VAR
BEGIN

REGION Network 1: Entradas Digitais
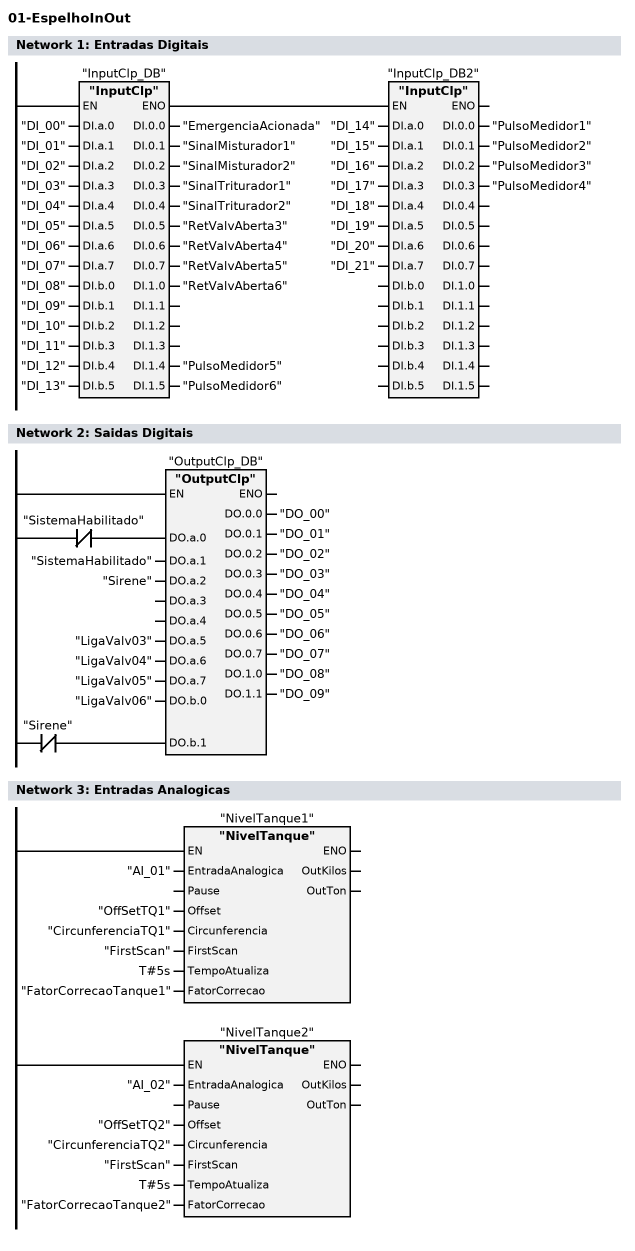
   RUNG wire#powerrail
      "InputClp_DB"("DI.a.0" := "DI_00", "DI.a.1" := "DI_01", "DI.a.2" := "DI_02", "DI.a.3" := "DI_03", "DI.a.4" := "DI_04", "DI.a.5" := "DI_05", "DI.a.6" := "DI_06", "DI.a.7" := "DI_07", "DI.b.0" := "DI_08", "DI.b.1" := "DI_09", "DI.b.2" := "DI_10", "DI.b.3" := "DI_11", "DI.b.4" := "DI_12", "DI.b.5" := "DI_13", "DI.0.0" => "EmergenciaAcionada", "DI.0.1" => "SinalMisturador1", "DI.0.2" => "SinalMisturador2", "DI.0.3" => "SinalTriturador1", "DI.0.4" => "SinalTriturador2", "DI.0.5" => "RetValvAberta3", "DI.0.6" => "RetValvAberta4", "DI.0.7" => "RetValvAberta5", "DI.1.0" => "RetValvAberta6", "DI.1.1" =>, "DI.1.2" =>, "DI.1.3" =>, "DI.1.4" => "PulsoMedidor5", "DI.1.5" => "PulsoMedidor6")
      "InputClp_DB2"("DI.a.0" := "DI_14", "DI.a.1" := "DI_15", "DI.a.2" := "DI_16", "DI.a.3" := "DI_17", "DI.a.4" := "DI_18", "DI.a.5" := "DI_19", "DI.a.6" := "DI_20", "DI.a.7" := "DI_21", "DI.b.0" :=, "DI.b.1" :=, "DI.b.2" :=, "DI.b.3" :=, "DI.b.4" :=, "DI.b.5" :=, "DI.0.0" => "PulsoMedidor1", "DI.0.1" => "PulsoMedidor2", "DI.0.2" => "PulsoMedidor3", "DI.0.3" => "PulsoMedidor4", "DI.0.4" =>, "DI.0.5" =>, "DI.0.6" =>, "DI.0.7" =>, "DI.1.0" =>, "DI.1.1" =>, "DI.1.2" =>, "DI.1.3" =>, "DI.1.4" =>, "DI.1.5" =>)
   END_RUNG
   // the same network as SCL:
   "InputClp_DB"("DI.a.0" := "DI_00",   // "InputClp"
                 "DI.a.1" := "DI_01",
                 "DI.a.2" := "DI_02",
                 "DI.a.3" := "DI_03",
                 "DI.a.4" := "DI_04",
                 "DI.a.5" := "DI_05",
                 "DI.a.6" := "DI_06",
                 "DI.a.7" := "DI_07",
                 "DI.b.0" := "DI_08",
                 "DI.b.1" := "DI_09",
                 "DI.b.2" := "DI_10",
                 "DI.b.3" := "DI_11",
                 "DI.b.4" := "DI_12",
                 "DI.b.5" := "DI_13",
                 "DI.0.0" => "EmergenciaAcionada",
                 "DI.0.1" => "SinalMisturador1",
                 "DI.0.2" => "SinalMisturador2",
                 "DI.0.3" => "SinalTriturador1",
                 "DI.0.4" => "SinalTriturador2",
                 "DI.0.5" => "RetValvAberta3",
                 "DI.0.6" => "RetValvAberta4",
                 "DI.0.7" => "RetValvAberta5",
                 "DI.1.0" => "RetValvAberta6",
                 "DI.1.4" => "PulsoMedidor5",
                 "DI.1.5" => "PulsoMedidor6",
                 ENO => #_w1);
   IF #_w1 THEN
       "InputClp_DB2"("DI.a.0" := "DI_14",   // "InputClp"
                      "DI.a.1" := "DI_15",
                      "DI.a.2" := "DI_16",
                      "DI.a.3" := "DI_17",
                      "DI.a.4" := "DI_18",
                      "DI.a.5" := "DI_19",
                      "DI.a.6" := "DI_20",
                      "DI.a.7" := "DI_21",
                      "DI.0.0" => "PulsoMedidor1",
                      "DI.0.1" => "PulsoMedidor2",
                      "DI.0.2" => "PulsoMedidor3",
                      "DI.0.3" => "PulsoMedidor4");
   END_IF;
END_REGION

REGION Network 2: Saidas Digitais
   RUNG wire#powerrail
      "OutputClp_DB"("DO.a.0" := wire#w1, "DO.b.1" := wire#w2, "DO.a.1" := "SistemaHabilitado", "DO.a.2" := "Sirene", "DO.a.3" :=, "DO.a.4" :=, "DO.a.5" := "LigaValv03", "DO.a.6" := "LigaValv04", "DO.a.7" := "LigaValv05", "DO.b.0" := "LigaValv06", "DO.0.0" => "DO_00", "DO.0.1" => "DO_01", "DO.0.2" => "DO_02", "DO.0.3" => "DO_03", "DO.0.4" => "DO_04", "DO.0.5" => "DO_05", "DO.0.6" => "DO_06", "DO.0.7" => "DO_07", "DO.1.0" => "DO_08", "DO.1.1" => "DO_09")
   END_RUNG
   RUNG wire#powerrail
      I_Contact( "SistemaHabilitado" )
   END_RUNG wire#w1
   RUNG wire#powerrail
      I_Contact( "Sirene" )
   END_RUNG wire#w2
   // the same network as SCL:
   "OutputClp_DB"("DO.a.0" := NOT "SistemaHabilitado",   // "OutputClp"
                  "DO.a.1" := "SistemaHabilitado",
                  "DO.a.2" := "Sirene",
                  "DO.a.5" := "LigaValv03",
                  "DO.a.6" := "LigaValv04",
                  "DO.a.7" := "LigaValv05",
                  "DO.b.0" := "LigaValv06",
                  "DO.b.1" := NOT "Sirene",
                  "DO.0.0" => "DO_00",
                  "DO.0.1" => "DO_01",
                  "DO.0.2" => "DO_02",
                  "DO.0.3" => "DO_03",
                  "DO.0.4" => "DO_04",
                  "DO.0.5" => "DO_05",
                  "DO.0.6" => "DO_06",
                  "DO.0.7" => "DO_07",
                  "DO.1.0" => "DO_08",
                  "DO.1.1" => "DO_09");
END_REGION

REGION Network 3: Entradas Analogicas
   RUNG wire#powerrail
      "NivelTanque1"(EntradaAnalogica := "AI_01", Pause :=, Offset := "OffSetTQ1", Circunferencia := "CircunferenciaTQ1", FirstScan := "FirstScan", TempoAtualiza := T#5s, FatorCorrecao := "FatorCorrecaoTanque1", OutKilos =>, OutTon =>)
   END_RUNG
   RUNG wire#powerrail
      "NivelTanque2"(EntradaAnalogica := "AI_02", Pause :=, Offset := "OffSetTQ2", Circunferencia := "CircunferenciaTQ2", FirstScan := "FirstScan", TempoAtualiza := T#5s, FatorCorrecao := "FatorCorrecaoTanque2", OutKilos =>, OutTon =>)
   END_RUNG
   // the same network as SCL:
   "NivelTanque1"(EntradaAnalogica := "AI_01",   // "NivelTanque"
                  Offset := "OffSetTQ1",
                  Circunferencia := "CircunferenciaTQ1",
                  FirstScan := "FirstScan",
                  TempoAtualiza := T#5s,
                  FatorCorrecao := "FatorCorrecaoTanque1");
   "NivelTanque2"(EntradaAnalogica := "AI_02",   // "NivelTanque"
                  Offset := "OffSetTQ2",
                  Circunferencia := "CircunferenciaTQ2",
                  FirstScan := "FirstScan",
                  TempoAtualiza := T#5s,
                  FatorCorrecao := "FatorCorrecaoTanque2");
END_REGION
END_ORGANIZATION_BLOCK

ORGANIZATION_BLOCK "02-Dosagem"   // OB124, LAD, ProgramCycle
TITLE = "Main Program Sweep (Cycle)"
{ S7_Optimized_Access := 'TRUE' }
VERSION : 0.1
   VAR_INPUT
      Initial_Call : Bool;   // Initial call of this OB
      Remanence : Bool;   // =True, if remanent data are available
   END_VAR
   VAR_TEMP   // added for the SCL form of the ladder/FBD networks
      _w1 : Bool;
      _w2 : Bool;
   END_VAR
BEGIN

REGION Network 1: Bomba 1 GamaX Triturador 1 Guardipet
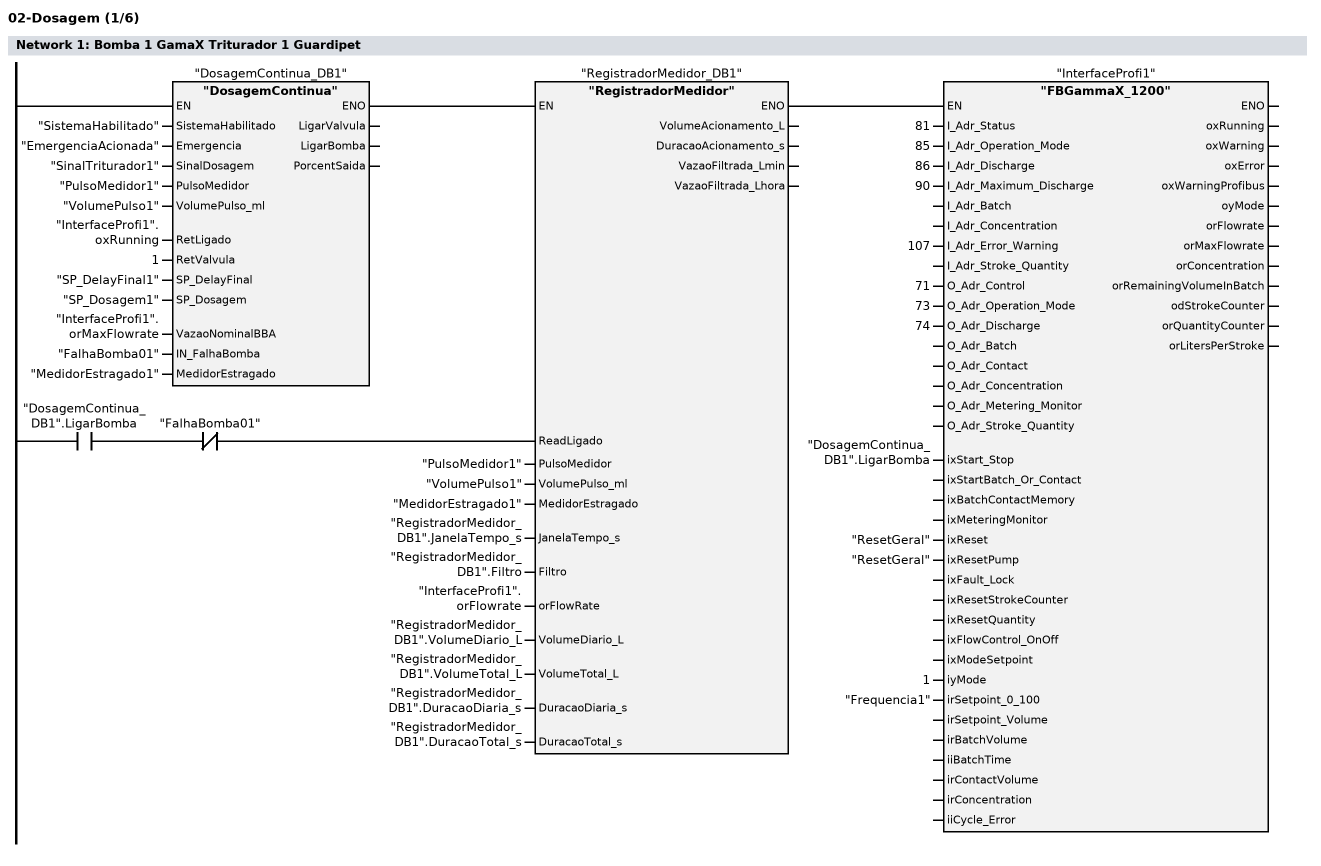
   RUNG wire#powerrail
      "DosagemContinua_DB1"(SistemaHabilitado := "SistemaHabilitado", Emergencia := "EmergenciaAcionada", SinalDosagem := "SinalTriturador1", PulsoMedidor := "PulsoMedidor1", VolumePulso_ml := "VolumePulso1", RetLigado := "InterfaceProfi1".oxRunning, RetValvula := 1, SP_DelayFinal := "SP_DelayFinal1", SP_Dosagem := "SP_Dosagem1", VazaoNominalBBA := "InterfaceProfi1".orMaxFlowrate, IN_FalhaBomba := "FalhaBomba01", MedidorEstragado := "MedidorEstragado1", LigarValvula =>, LigarBomba =>, PorcentSaida =>)
      "RegistradorMedidor_DB1"(ReadLigado := wire#w1, PulsoMedidor := "PulsoMedidor1", VolumePulso_ml := "VolumePulso1", MedidorEstragado := "MedidorEstragado1", JanelaTempo_s := "RegistradorMedidor_DB1".JanelaTempo_s, Filtro := "RegistradorMedidor_DB1".Filtro, orFlowRate := "InterfaceProfi1".orFlowrate, VolumeDiario_L := "RegistradorMedidor_DB1".VolumeDiario_L, VolumeTotal_L := "RegistradorMedidor_DB1".VolumeTotal_L, DuracaoDiaria_s := "RegistradorMedidor_DB1".DuracaoDiaria_s, DuracaoTotal_s := "RegistradorMedidor_DB1".DuracaoTotal_s, VolumeAcionamento_L =>, DuracaoAcionamento_s =>, VazaoFiltrada_Lmin =>, VazaoFiltrada_Lhora =>)
      "InterfaceProfi1"(I_Adr_Status := 81, I_Adr_Operation_Mode := 85, I_Adr_Discharge := 86, I_Adr_Maximum_Discharge := 90, I_Adr_Batch :=, I_Adr_Concentration :=, I_Adr_Error_Warning := 107, I_Adr_Stroke_Quantity :=, O_Adr_Control := 71, O_Adr_Operation_Mode := 73, O_Adr_Discharge := 74, O_Adr_Batch :=, O_Adr_Contact :=, O_Adr_Concentration :=, O_Adr_Metering_Monitor :=, O_Adr_Stroke_Quantity :=, ixStart_Stop := "DosagemContinua_DB1".LigarBomba, ixStartBatch_Or_Contact :=, ixBatchContactMemory :=, ixMeteringMonitor :=, ixReset := "ResetGeral", ixResetPump := "ResetGeral", ixFault_Lock :=, ixResetStrokeCounter :=, ixResetQuantity :=, ixFlowControl_OnOff :=, ixModeSetpoint :=, iyMode := 1, irSetpoint_0_100 := "Frequencia1", irSetpoint_Volume :=, irBatchVolume :=, iiBatchTime :=, irContactVolume :=, irConcentration :=, iiCycle_Error :=, oxRunning =>, oxWarning =>, oxError =>, oxWarningProfibus =>, oyMode =>, orFlowrate =>, orMaxFlowrate =>, orConcentration =>, orRemainingVolumeInBatch =>, odStrokeCounter =>, orQuantityCounter =>, orLitersPerStroke =>)
   END_RUNG
   RUNG wire#powerrail
      Contact( "DosagemContinua_DB1".LigarBomba )
      I_Contact( "FalhaBomba01" )
   END_RUNG wire#w1
   // the same network as SCL:
   "DosagemContinua_DB1"(SistemaHabilitado := "SistemaHabilitado",   // "DosagemContinua"
                         Emergencia := "EmergenciaAcionada",
                         SinalDosagem := "SinalTriturador1",
                         PulsoMedidor := "PulsoMedidor1",
                         VolumePulso_ml := "VolumePulso1",
                         RetLigado := "InterfaceProfi1".oxRunning,
                         RetValvula := 1,
                         SP_DelayFinal := "SP_DelayFinal1",
                         SP_Dosagem := "SP_Dosagem1",
                         VazaoNominalBBA := "InterfaceProfi1".orMaxFlowrate,
                         IN_FalhaBomba := "FalhaBomba01",
                         MedidorEstragado := "MedidorEstragado1",
                         ENO => #_w1);
   "RegistradorMedidor_DB1"(EN := #_w1,   // "RegistradorMedidor"
                           ReadLigado := "DosagemContinua_DB1".LigarBomba AND NOT "FalhaBomba01",
                           PulsoMedidor := "PulsoMedidor1",
                           VolumePulso_ml := "VolumePulso1",
                           MedidorEstragado := "MedidorEstragado1",
                           JanelaTempo_s := "RegistradorMedidor_DB1".JanelaTempo_s,
                           Filtro := "RegistradorMedidor_DB1".Filtro,
                           orFlowRate := "InterfaceProfi1".orFlowrate,
                           VolumeDiario_L := "RegistradorMedidor_DB1".VolumeDiario_L,
                           VolumeTotal_L := "RegistradorMedidor_DB1".VolumeTotal_L,
                           DuracaoDiaria_s := "RegistradorMedidor_DB1".DuracaoDiaria_s,
                           DuracaoTotal_s := "RegistradorMedidor_DB1".DuracaoTotal_s,
                           ENO => #_w2);
   IF #_w2 THEN
       "InterfaceProfi1"(I_Adr_Status := 81,   // "FBGammaX_1200"
                         I_Adr_Operation_Mode := 85,
                         I_Adr_Discharge := 86,
                         I_Adr_Maximum_Discharge := 90,
                         I_Adr_Error_Warning := 107,
                         O_Adr_Control := 71,
                         O_Adr_Operation_Mode := 73,
                         O_Adr_Discharge := 74,
                         ixStart_Stop := "DosagemContinua_DB1".LigarBomba,
                         ixReset := "ResetGeral",
                         ixResetPump := "ResetGeral",
                         iyMode := 1,
                         irSetpoint_0_100 := "Frequencia1");
   END_IF;
END_REGION

REGION Network 2: Bomba 2 GamaX Triturador 2 Guardipet
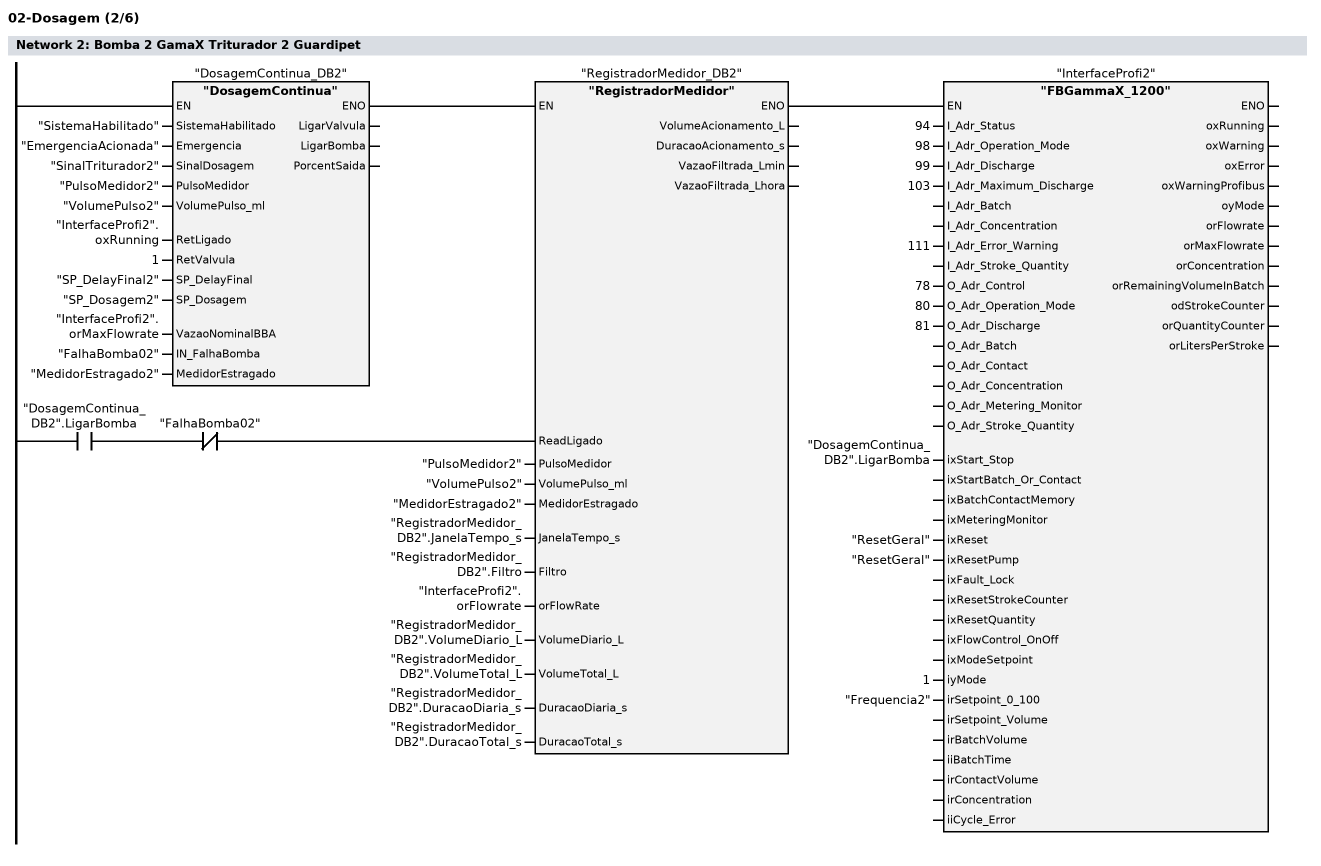
   RUNG wire#powerrail
      "DosagemContinua_DB2"(SistemaHabilitado := "SistemaHabilitado", Emergencia := "EmergenciaAcionada", SinalDosagem := "SinalTriturador2", PulsoMedidor := "PulsoMedidor2", VolumePulso_ml := "VolumePulso2", RetLigado := "InterfaceProfi2".oxRunning, RetValvula := 1, SP_DelayFinal := "SP_DelayFinal2", SP_Dosagem := "SP_Dosagem2", VazaoNominalBBA := "InterfaceProfi2".orMaxFlowrate, IN_FalhaBomba := "FalhaBomba02", MedidorEstragado := "MedidorEstragado2", LigarValvula =>, LigarBomba =>, PorcentSaida =>)
      "RegistradorMedidor_DB2"(ReadLigado := wire#w1, PulsoMedidor := "PulsoMedidor2", VolumePulso_ml := "VolumePulso2", MedidorEstragado := "MedidorEstragado2", JanelaTempo_s := "RegistradorMedidor_DB2".JanelaTempo_s, Filtro := "RegistradorMedidor_DB2".Filtro, orFlowRate := "InterfaceProfi2".orFlowrate, VolumeDiario_L := "RegistradorMedidor_DB2".VolumeDiario_L, VolumeTotal_L := "RegistradorMedidor_DB2".VolumeTotal_L, DuracaoDiaria_s := "RegistradorMedidor_DB2".DuracaoDiaria_s, DuracaoTotal_s := "RegistradorMedidor_DB2".DuracaoTotal_s, VolumeAcionamento_L =>, DuracaoAcionamento_s =>, VazaoFiltrada_Lmin =>, VazaoFiltrada_Lhora =>)
      "InterfaceProfi2"(I_Adr_Status := 94, I_Adr_Operation_Mode := 98, I_Adr_Discharge := 99, I_Adr_Maximum_Discharge := 103, I_Adr_Batch :=, I_Adr_Concentration :=, I_Adr_Error_Warning := 111, I_Adr_Stroke_Quantity :=, O_Adr_Control := 78, O_Adr_Operation_Mode := 80, O_Adr_Discharge := 81, O_Adr_Batch :=, O_Adr_Contact :=, O_Adr_Concentration :=, O_Adr_Metering_Monitor :=, O_Adr_Stroke_Quantity :=, ixStart_Stop := "DosagemContinua_DB2".LigarBomba, ixStartBatch_Or_Contact :=, ixBatchContactMemory :=, ixMeteringMonitor :=, ixReset := "ResetGeral", ixResetPump := "ResetGeral", ixFault_Lock :=, ixResetStrokeCounter :=, ixResetQuantity :=, ixFlowControl_OnOff :=, ixModeSetpoint :=, iyMode := 1, irSetpoint_0_100 := "Frequencia2", irSetpoint_Volume :=, irBatchVolume :=, iiBatchTime :=, irContactVolume :=, irConcentration :=, iiCycle_Error :=, oxRunning =>, oxWarning =>, oxError =>, oxWarningProfibus =>, oyMode =>, orFlowrate =>, orMaxFlowrate =>, orConcentration =>, orRemainingVolumeInBatch =>, odStrokeCounter =>, orQuantityCounter =>, orLitersPerStroke =>)
   END_RUNG
   RUNG wire#powerrail
      Contact( "DosagemContinua_DB2".LigarBomba )
      I_Contact( "FalhaBomba02" )
   END_RUNG wire#w1
   // the same network as SCL:
   "DosagemContinua_DB2"(SistemaHabilitado := "SistemaHabilitado",   // "DosagemContinua"
                         Emergencia := "EmergenciaAcionada",
                         SinalDosagem := "SinalTriturador2",
                         PulsoMedidor := "PulsoMedidor2",
                         VolumePulso_ml := "VolumePulso2",
                         RetLigado := "InterfaceProfi2".oxRunning,
                         RetValvula := 1,
                         SP_DelayFinal := "SP_DelayFinal2",
                         SP_Dosagem := "SP_Dosagem2",
                         VazaoNominalBBA := "InterfaceProfi2".orMaxFlowrate,
                         IN_FalhaBomba := "FalhaBomba02",
                         MedidorEstragado := "MedidorEstragado2",
                         ENO => #_w1);
   "RegistradorMedidor_DB2"(EN := #_w1,   // "RegistradorMedidor"
                           ReadLigado := "DosagemContinua_DB2".LigarBomba AND NOT "FalhaBomba02",
                           PulsoMedidor := "PulsoMedidor2",
                           VolumePulso_ml := "VolumePulso2",
                           MedidorEstragado := "MedidorEstragado2",
                           JanelaTempo_s := "RegistradorMedidor_DB2".JanelaTempo_s,
                           Filtro := "RegistradorMedidor_DB2".Filtro,
                           orFlowRate := "InterfaceProfi2".orFlowrate,
                           VolumeDiario_L := "RegistradorMedidor_DB2".VolumeDiario_L,
                           VolumeTotal_L := "RegistradorMedidor_DB2".VolumeTotal_L,
                           DuracaoDiaria_s := "RegistradorMedidor_DB2".DuracaoDiaria_s,
                           DuracaoTotal_s := "RegistradorMedidor_DB2".DuracaoTotal_s,
                           ENO => #_w2);
   IF #_w2 THEN
       "InterfaceProfi2"(I_Adr_Status := 94,   // "FBGammaX_1200"
                         I_Adr_Operation_Mode := 98,
                         I_Adr_Discharge := 99,
                         I_Adr_Maximum_Discharge := 103,
                         I_Adr_Error_Warning := 111,
                         O_Adr_Control := 78,
                         O_Adr_Operation_Mode := 80,
                         O_Adr_Discharge := 81,
                         ixStart_Stop := "DosagemContinua_DB2".LigarBomba,
                         ixReset := "ResetGeral",
                         ixResetPump := "ResetGeral",
                         iyMode := 1,
                         irSetpoint_0_100 := "Frequencia2");
   END_IF;
END_REGION

REGION Network 3: Bomba 3 GamaX Misturador 1 Guardipet
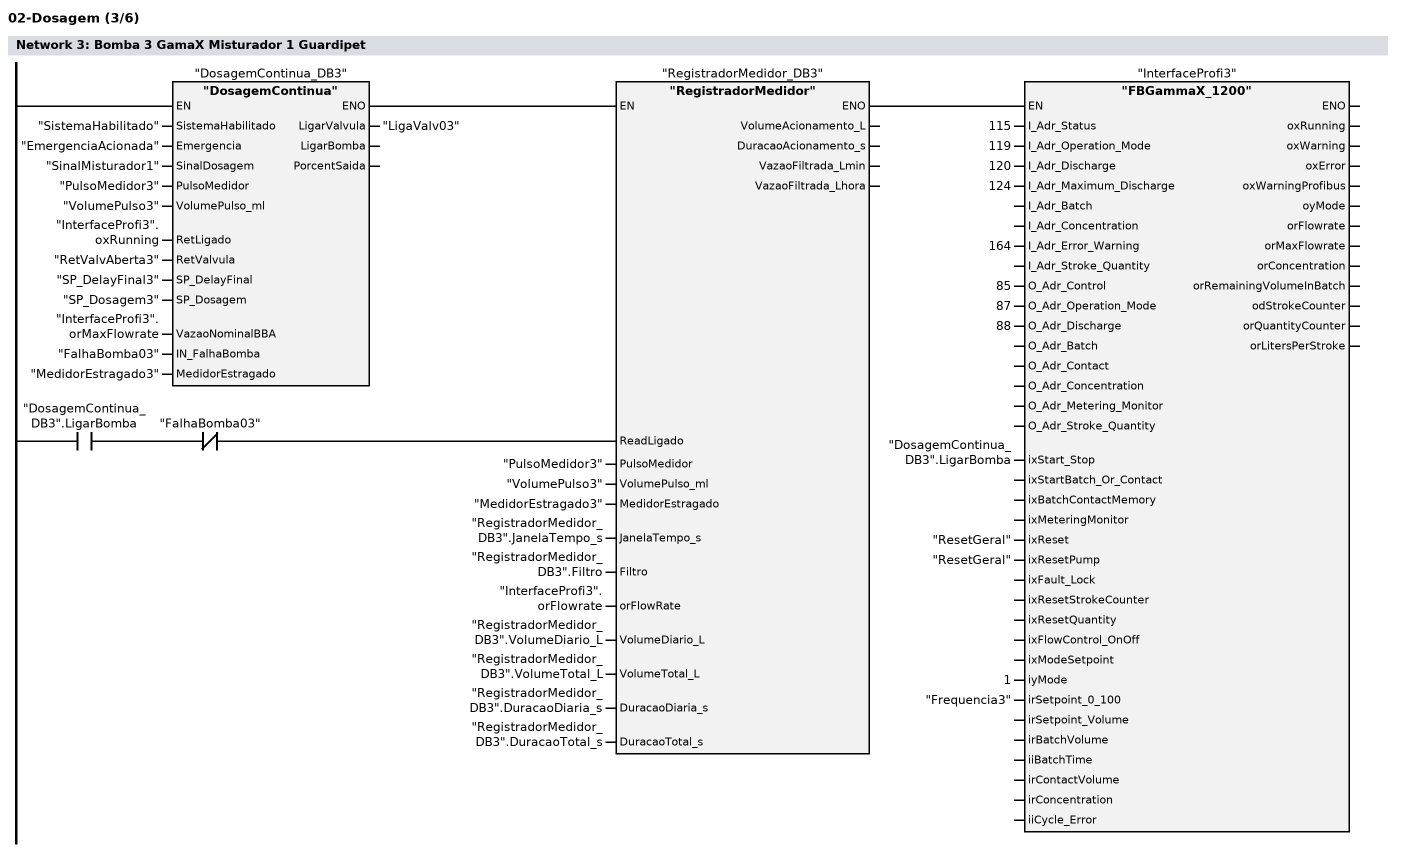
   RUNG wire#powerrail
      "DosagemContinua_DB3"(SistemaHabilitado := "SistemaHabilitado", Emergencia := "EmergenciaAcionada", SinalDosagem := "SinalMisturador1", PulsoMedidor := "PulsoMedidor3", VolumePulso_ml := "VolumePulso3", RetLigado := "InterfaceProfi3".oxRunning, RetValvula := "RetValvAberta3", SP_DelayFinal := "SP_DelayFinal3", SP_Dosagem := "SP_Dosagem3", VazaoNominalBBA := "InterfaceProfi3".orMaxFlowrate, IN_FalhaBomba := "FalhaBomba03", MedidorEstragado := "MedidorEstragado3", LigarValvula => "LigaValv03", LigarBomba =>, PorcentSaida =>)
      "RegistradorMedidor_DB3"(ReadLigado := wire#w1, PulsoMedidor := "PulsoMedidor3", VolumePulso_ml := "VolumePulso3", MedidorEstragado := "MedidorEstragado3", JanelaTempo_s := "RegistradorMedidor_DB3".JanelaTempo_s, Filtro := "RegistradorMedidor_DB3".Filtro, orFlowRate := "InterfaceProfi3".orFlowrate, VolumeDiario_L := "RegistradorMedidor_DB3".VolumeDiario_L, VolumeTotal_L := "RegistradorMedidor_DB3".VolumeTotal_L, DuracaoDiaria_s := "RegistradorMedidor_DB3".DuracaoDiaria_s, DuracaoTotal_s := "RegistradorMedidor_DB3".DuracaoTotal_s, VolumeAcionamento_L =>, DuracaoAcionamento_s =>, VazaoFiltrada_Lmin =>, VazaoFiltrada_Lhora =>)
      "InterfaceProfi3"(I_Adr_Status := 115, I_Adr_Operation_Mode := 119, I_Adr_Discharge := 120, I_Adr_Maximum_Discharge := 124, I_Adr_Batch :=, I_Adr_Concentration :=, I_Adr_Error_Warning := 164, I_Adr_Stroke_Quantity :=, O_Adr_Control := 85, O_Adr_Operation_Mode := 87, O_Adr_Discharge := 88, O_Adr_Batch :=, O_Adr_Contact :=, O_Adr_Concentration :=, O_Adr_Metering_Monitor :=, O_Adr_Stroke_Quantity :=, ixStart_Stop := "DosagemContinua_DB3".LigarBomba, ixStartBatch_Or_Contact :=, ixBatchContactMemory :=, ixMeteringMonitor :=, ixReset := "ResetGeral", ixResetPump := "ResetGeral", ixFault_Lock :=, ixResetStrokeCounter :=, ixResetQuantity :=, ixFlowControl_OnOff :=, ixModeSetpoint :=, iyMode := 1, irSetpoint_0_100 := "Frequencia3", irSetpoint_Volume :=, irBatchVolume :=, iiBatchTime :=, irContactVolume :=, irConcentration :=, iiCycle_Error :=, oxRunning =>, oxWarning =>, oxError =>, oxWarningProfibus =>, oyMode =>, orFlowrate =>, orMaxFlowrate =>, orConcentration =>, orRemainingVolumeInBatch =>, odStrokeCounter =>, orQuantityCounter =>, orLitersPerStroke =>)
   END_RUNG
   RUNG wire#powerrail
      Contact( "DosagemContinua_DB3".LigarBomba )
      I_Contact( "FalhaBomba03" )
   END_RUNG wire#w1
   // the same network as SCL:
   "DosagemContinua_DB3"(SistemaHabilitado := "SistemaHabilitado",   // "DosagemContinua"
                         Emergencia := "EmergenciaAcionada",
                         SinalDosagem := "SinalMisturador1",
                         PulsoMedidor := "PulsoMedidor3",
                         VolumePulso_ml := "VolumePulso3",
                         RetLigado := "InterfaceProfi3".oxRunning,
                         RetValvula := "RetValvAberta3",
                         SP_DelayFinal := "SP_DelayFinal3",
                         SP_Dosagem := "SP_Dosagem3",
                         VazaoNominalBBA := "InterfaceProfi3".orMaxFlowrate,
                         IN_FalhaBomba := "FalhaBomba03",
                         MedidorEstragado := "MedidorEstragado3",
                         LigarValvula => "LigaValv03",
                         ENO => #_w1);
   "RegistradorMedidor_DB3"(EN := #_w1,   // "RegistradorMedidor"
                           ReadLigado := "DosagemContinua_DB3".LigarBomba AND NOT "FalhaBomba03",
                           PulsoMedidor := "PulsoMedidor3",
                           VolumePulso_ml := "VolumePulso3",
                           MedidorEstragado := "MedidorEstragado3",
                           JanelaTempo_s := "RegistradorMedidor_DB3".JanelaTempo_s,
                           Filtro := "RegistradorMedidor_DB3".Filtro,
                           orFlowRate := "InterfaceProfi3".orFlowrate,
                           VolumeDiario_L := "RegistradorMedidor_DB3".VolumeDiario_L,
                           VolumeTotal_L := "RegistradorMedidor_DB3".VolumeTotal_L,
                           DuracaoDiaria_s := "RegistradorMedidor_DB3".DuracaoDiaria_s,
                           DuracaoTotal_s := "RegistradorMedidor_DB3".DuracaoTotal_s,
                           ENO => #_w2);
   IF #_w2 THEN
       "InterfaceProfi3"(I_Adr_Status := 115,   // "FBGammaX_1200"
                         I_Adr_Operation_Mode := 119,
                         I_Adr_Discharge := 120,
                         I_Adr_Maximum_Discharge := 124,
                         I_Adr_Error_Warning := 164,
                         O_Adr_Control := 85,
                         O_Adr_Operation_Mode := 87,
                         O_Adr_Discharge := 88,
                         ixStart_Stop := "DosagemContinua_DB3".LigarBomba,
                         ixReset := "ResetGeral",
                         ixResetPump := "ResetGeral",
                         iyMode := 1,
                         irSetpoint_0_100 := "Frequencia3");
   END_IF;
END_REGION

REGION Network 4: Bomba 4 GamaX Misturador 2 Guardipet
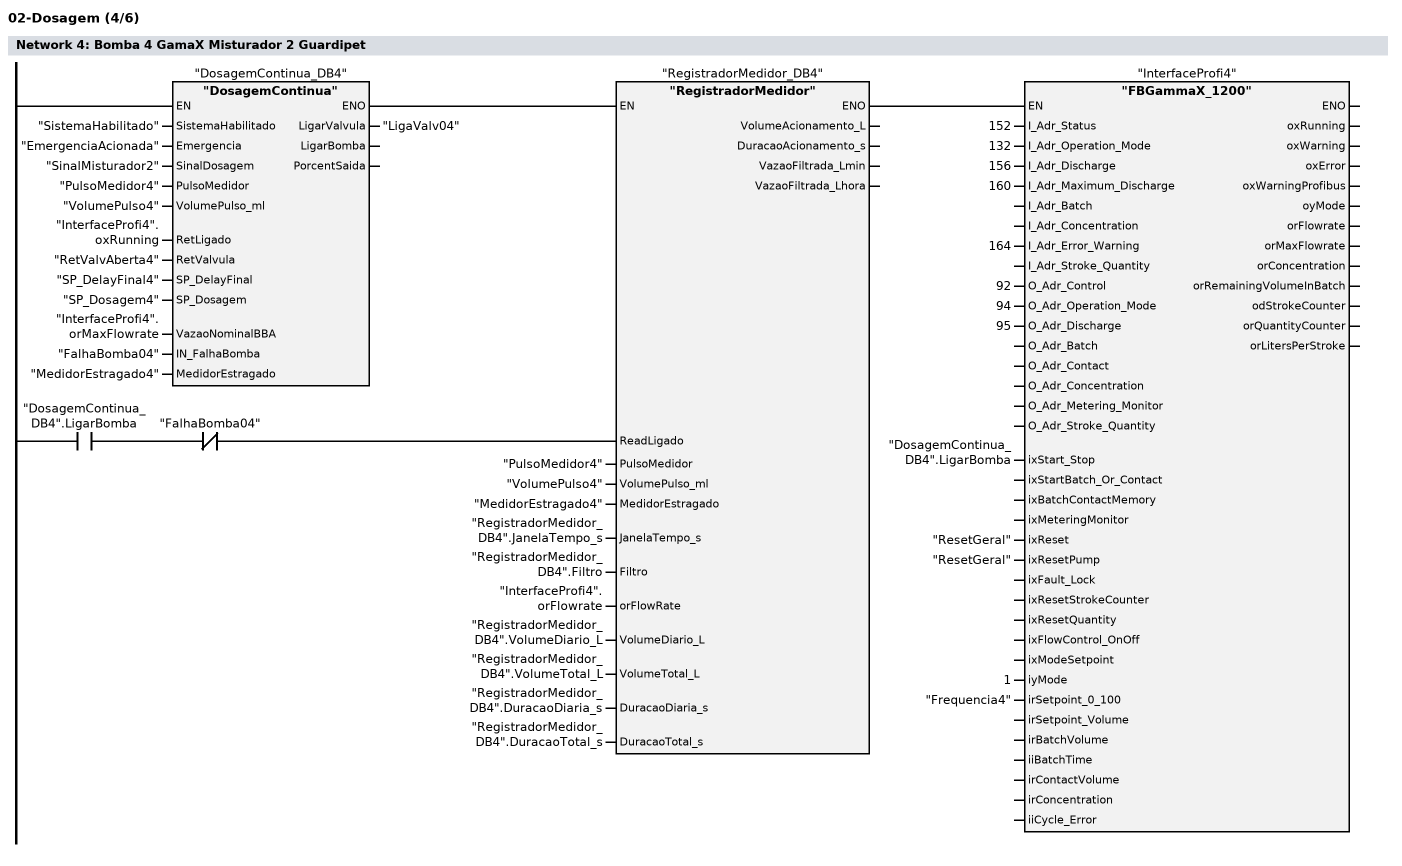
   RUNG wire#powerrail
      "DosagemContinua_DB4"(SistemaHabilitado := "SistemaHabilitado", Emergencia := "EmergenciaAcionada", SinalDosagem := "SinalMisturador2", PulsoMedidor := "PulsoMedidor4", VolumePulso_ml := "VolumePulso4", RetLigado := "InterfaceProfi4".oxRunning, RetValvula := "RetValvAberta4", SP_DelayFinal := "SP_DelayFinal4", SP_Dosagem := "SP_Dosagem4", VazaoNominalBBA := "InterfaceProfi4".orMaxFlowrate, IN_FalhaBomba := "FalhaBomba04", MedidorEstragado := "MedidorEstragado4", LigarValvula => "LigaValv04", LigarBomba =>, PorcentSaida =>)
      "RegistradorMedidor_DB4"(ReadLigado := wire#w1, PulsoMedidor := "PulsoMedidor4", VolumePulso_ml := "VolumePulso4", MedidorEstragado := "MedidorEstragado4", JanelaTempo_s := "RegistradorMedidor_DB4".JanelaTempo_s, Filtro := "RegistradorMedidor_DB4".Filtro, orFlowRate := "InterfaceProfi4".orFlowrate, VolumeDiario_L := "RegistradorMedidor_DB4".VolumeDiario_L, VolumeTotal_L := "RegistradorMedidor_DB4".VolumeTotal_L, DuracaoDiaria_s := "RegistradorMedidor_DB4".DuracaoDiaria_s, DuracaoTotal_s := "RegistradorMedidor_DB4".DuracaoTotal_s, VolumeAcionamento_L =>, DuracaoAcionamento_s =>, VazaoFiltrada_Lmin =>, VazaoFiltrada_Lhora =>)
      "InterfaceProfi4"(I_Adr_Status := 152, I_Adr_Operation_Mode := 132, I_Adr_Discharge := 156, I_Adr_Maximum_Discharge := 160, I_Adr_Batch :=, I_Adr_Concentration :=, I_Adr_Error_Warning := 164, I_Adr_Stroke_Quantity :=, O_Adr_Control := 92, O_Adr_Operation_Mode := 94, O_Adr_Discharge := 95, O_Adr_Batch :=, O_Adr_Contact :=, O_Adr_Concentration :=, O_Adr_Metering_Monitor :=, O_Adr_Stroke_Quantity :=, ixStart_Stop := "DosagemContinua_DB4".LigarBomba, ixStartBatch_Or_Contact :=, ixBatchContactMemory :=, ixMeteringMonitor :=, ixReset := "ResetGeral", ixResetPump := "ResetGeral", ixFault_Lock :=, ixResetStrokeCounter :=, ixResetQuantity :=, ixFlowControl_OnOff :=, ixModeSetpoint :=, iyMode := 1, irSetpoint_0_100 := "Frequencia4", irSetpoint_Volume :=, irBatchVolume :=, iiBatchTime :=, irContactVolume :=, irConcentration :=, iiCycle_Error :=, oxRunning =>, oxWarning =>, oxError =>, oxWarningProfibus =>, oyMode =>, orFlowrate =>, orMaxFlowrate =>, orConcentration =>, orRemainingVolumeInBatch =>, odStrokeCounter =>, orQuantityCounter =>, orLitersPerStroke =>)
   END_RUNG
   RUNG wire#powerrail
      Contact( "DosagemContinua_DB4".LigarBomba )
      I_Contact( "FalhaBomba04" )
   END_RUNG wire#w1
   // the same network as SCL:
   "DosagemContinua_DB4"(SistemaHabilitado := "SistemaHabilitado",   // "DosagemContinua"
                         Emergencia := "EmergenciaAcionada",
                         SinalDosagem := "SinalMisturador2",
                         PulsoMedidor := "PulsoMedidor4",
                         VolumePulso_ml := "VolumePulso4",
                         RetLigado := "InterfaceProfi4".oxRunning,
                         RetValvula := "RetValvAberta4",
                         SP_DelayFinal := "SP_DelayFinal4",
                         SP_Dosagem := "SP_Dosagem4",
                         VazaoNominalBBA := "InterfaceProfi4".orMaxFlowrate,
                         IN_FalhaBomba := "FalhaBomba04",
                         MedidorEstragado := "MedidorEstragado4",
                         LigarValvula => "LigaValv04",
                         ENO => #_w1);
   "RegistradorMedidor_DB4"(EN := #_w1,   // "RegistradorMedidor"
                           ReadLigado := "DosagemContinua_DB4".LigarBomba AND NOT "FalhaBomba04",
                           PulsoMedidor := "PulsoMedidor4",
                           VolumePulso_ml := "VolumePulso4",
                           MedidorEstragado := "MedidorEstragado4",
                           JanelaTempo_s := "RegistradorMedidor_DB4".JanelaTempo_s,
                           Filtro := "RegistradorMedidor_DB4".Filtro,
                           orFlowRate := "InterfaceProfi4".orFlowrate,
                           VolumeDiario_L := "RegistradorMedidor_DB4".VolumeDiario_L,
                           VolumeTotal_L := "RegistradorMedidor_DB4".VolumeTotal_L,
                           DuracaoDiaria_s := "RegistradorMedidor_DB4".DuracaoDiaria_s,
                           DuracaoTotal_s := "RegistradorMedidor_DB4".DuracaoTotal_s,
                           ENO => #_w2);
   IF #_w2 THEN
       "InterfaceProfi4"(I_Adr_Status := 152,   // "FBGammaX_1200"
                         I_Adr_Operation_Mode := 132,
                         I_Adr_Discharge := 156,
                         I_Adr_Maximum_Discharge := 160,
                         I_Adr_Error_Warning := 164,
                         O_Adr_Control := 92,
                         O_Adr_Operation_Mode := 94,
                         O_Adr_Discharge := 95,
                         ixStart_Stop := "DosagemContinua_DB4".LigarBomba,
                         ixReset := "ResetGeral",
                         ixResetPump := "ResetGeral",
                         iyMode := 1,
                         irSetpoint_0_100 := "Frequencia4");
   END_IF;
END_REGION

REGION Network 5: Bomba 5 GamaX Misturador 1 Bactonew
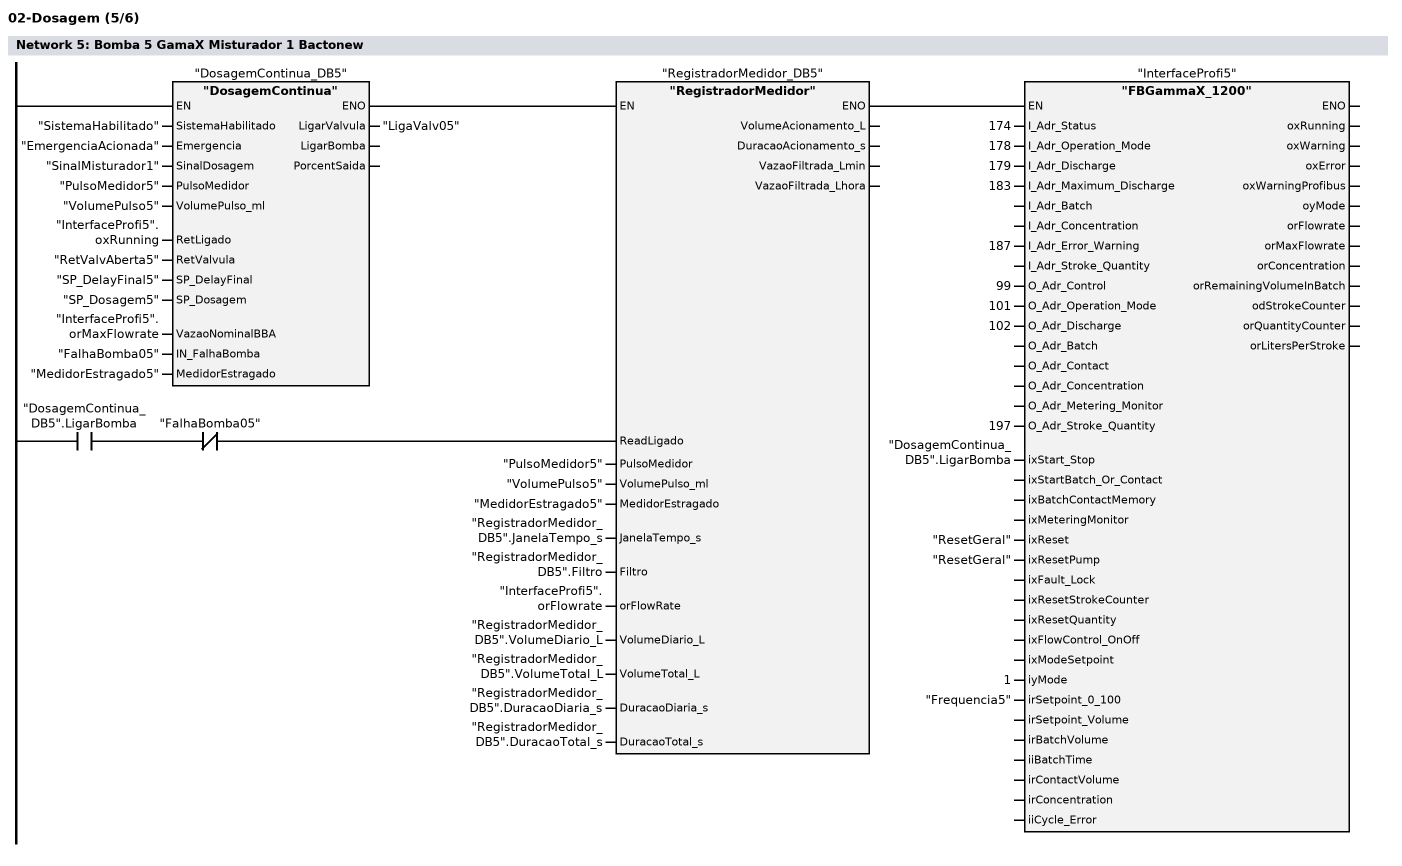
   RUNG wire#powerrail
      "DosagemContinua_DB5"(SistemaHabilitado := "SistemaHabilitado", Emergencia := "EmergenciaAcionada", SinalDosagem := "SinalMisturador1", PulsoMedidor := "PulsoMedidor5", VolumePulso_ml := "VolumePulso5", RetLigado := "InterfaceProfi5".oxRunning, RetValvula := "RetValvAberta5", SP_DelayFinal := "SP_DelayFinal5", SP_Dosagem := "SP_Dosagem5", VazaoNominalBBA := "InterfaceProfi5".orMaxFlowrate, IN_FalhaBomba := "FalhaBomba05", MedidorEstragado := "MedidorEstragado5", LigarValvula => "LigaValv05", LigarBomba =>, PorcentSaida =>)
      "RegistradorMedidor_DB5"(ReadLigado := wire#w1, PulsoMedidor := "PulsoMedidor5", VolumePulso_ml := "VolumePulso5", MedidorEstragado := "MedidorEstragado5", JanelaTempo_s := "RegistradorMedidor_DB5".JanelaTempo_s, Filtro := "RegistradorMedidor_DB5".Filtro, orFlowRate := "InterfaceProfi5".orFlowrate, VolumeDiario_L := "RegistradorMedidor_DB5".VolumeDiario_L, VolumeTotal_L := "RegistradorMedidor_DB5".VolumeTotal_L, DuracaoDiaria_s := "RegistradorMedidor_DB5".DuracaoDiaria_s, DuracaoTotal_s := "RegistradorMedidor_DB5".DuracaoTotal_s, VolumeAcionamento_L =>, DuracaoAcionamento_s =>, VazaoFiltrada_Lmin =>, VazaoFiltrada_Lhora =>)
      "InterfaceProfi5"(I_Adr_Status := 174, I_Adr_Operation_Mode := 178, I_Adr_Discharge := 179, I_Adr_Maximum_Discharge := 183, I_Adr_Batch :=, I_Adr_Concentration :=, I_Adr_Error_Warning := 187, I_Adr_Stroke_Quantity :=, O_Adr_Control := 99, O_Adr_Operation_Mode := 101, O_Adr_Discharge := 102, O_Adr_Batch :=, O_Adr_Contact :=, O_Adr_Concentration :=, O_Adr_Metering_Monitor :=, O_Adr_Stroke_Quantity := 197, ixStart_Stop := "DosagemContinua_DB5".LigarBomba, ixStartBatch_Or_Contact :=, ixBatchContactMemory :=, ixMeteringMonitor :=, ixReset := "ResetGeral", ixResetPump := "ResetGeral", ixFault_Lock :=, ixResetStrokeCounter :=, ixResetQuantity :=, ixFlowControl_OnOff :=, ixModeSetpoint :=, iyMode := 1, irSetpoint_0_100 := "Frequencia5", irSetpoint_Volume :=, irBatchVolume :=, iiBatchTime :=, irContactVolume :=, irConcentration :=, iiCycle_Error :=, oxRunning =>, oxWarning =>, oxError =>, oxWarningProfibus =>, oyMode =>, orFlowrate =>, orMaxFlowrate =>, orConcentration =>, orRemainingVolumeInBatch =>, odStrokeCounter =>, orQuantityCounter =>, orLitersPerStroke =>)
   END_RUNG
   RUNG wire#powerrail
      Contact( "DosagemContinua_DB5".LigarBomba )
      I_Contact( "FalhaBomba05" )
   END_RUNG wire#w1
   // the same network as SCL:
   "DosagemContinua_DB5"(SistemaHabilitado := "SistemaHabilitado",   // "DosagemContinua"
                         Emergencia := "EmergenciaAcionada",
                         SinalDosagem := "SinalMisturador1",
                         PulsoMedidor := "PulsoMedidor5",
                         VolumePulso_ml := "VolumePulso5",
                         RetLigado := "InterfaceProfi5".oxRunning,
                         RetValvula := "RetValvAberta5",
                         SP_DelayFinal := "SP_DelayFinal5",
                         SP_Dosagem := "SP_Dosagem5",
                         VazaoNominalBBA := "InterfaceProfi5".orMaxFlowrate,
                         IN_FalhaBomba := "FalhaBomba05",
                         MedidorEstragado := "MedidorEstragado5",
                         LigarValvula => "LigaValv05",
                         ENO => #_w1);
   "RegistradorMedidor_DB5"(EN := #_w1,   // "RegistradorMedidor"
                           ReadLigado := "DosagemContinua_DB5".LigarBomba AND NOT "FalhaBomba05",
                           PulsoMedidor := "PulsoMedidor5",
                           VolumePulso_ml := "VolumePulso5",
                           MedidorEstragado := "MedidorEstragado5",
                           JanelaTempo_s := "RegistradorMedidor_DB5".JanelaTempo_s,
                           Filtro := "RegistradorMedidor_DB5".Filtro,
                           orFlowRate := "InterfaceProfi5".orFlowrate,
                           VolumeDiario_L := "RegistradorMedidor_DB5".VolumeDiario_L,
                           VolumeTotal_L := "RegistradorMedidor_DB5".VolumeTotal_L,
                           DuracaoDiaria_s := "RegistradorMedidor_DB5".DuracaoDiaria_s,
                           DuracaoTotal_s := "RegistradorMedidor_DB5".DuracaoTotal_s,
                           ENO => #_w2);
   IF #_w2 THEN
       "InterfaceProfi5"(I_Adr_Status := 174,   // "FBGammaX_1200"
                         I_Adr_Operation_Mode := 178,
                         I_Adr_Discharge := 179,
                         I_Adr_Maximum_Discharge := 183,
                         I_Adr_Error_Warning := 187,
                         O_Adr_Control := 99,
                         O_Adr_Operation_Mode := 101,
                         O_Adr_Discharge := 102,
                         O_Adr_Stroke_Quantity := 197,
                         ixStart_Stop := "DosagemContinua_DB5".LigarBomba,
                         ixReset := "ResetGeral",
                         ixResetPump := "ResetGeral",
                         iyMode := 1,
                         irSetpoint_0_100 := "Frequencia5");
   END_IF;
END_REGION

REGION Network 6: Bomba 6 GamaX Misturador 2 Bactonew
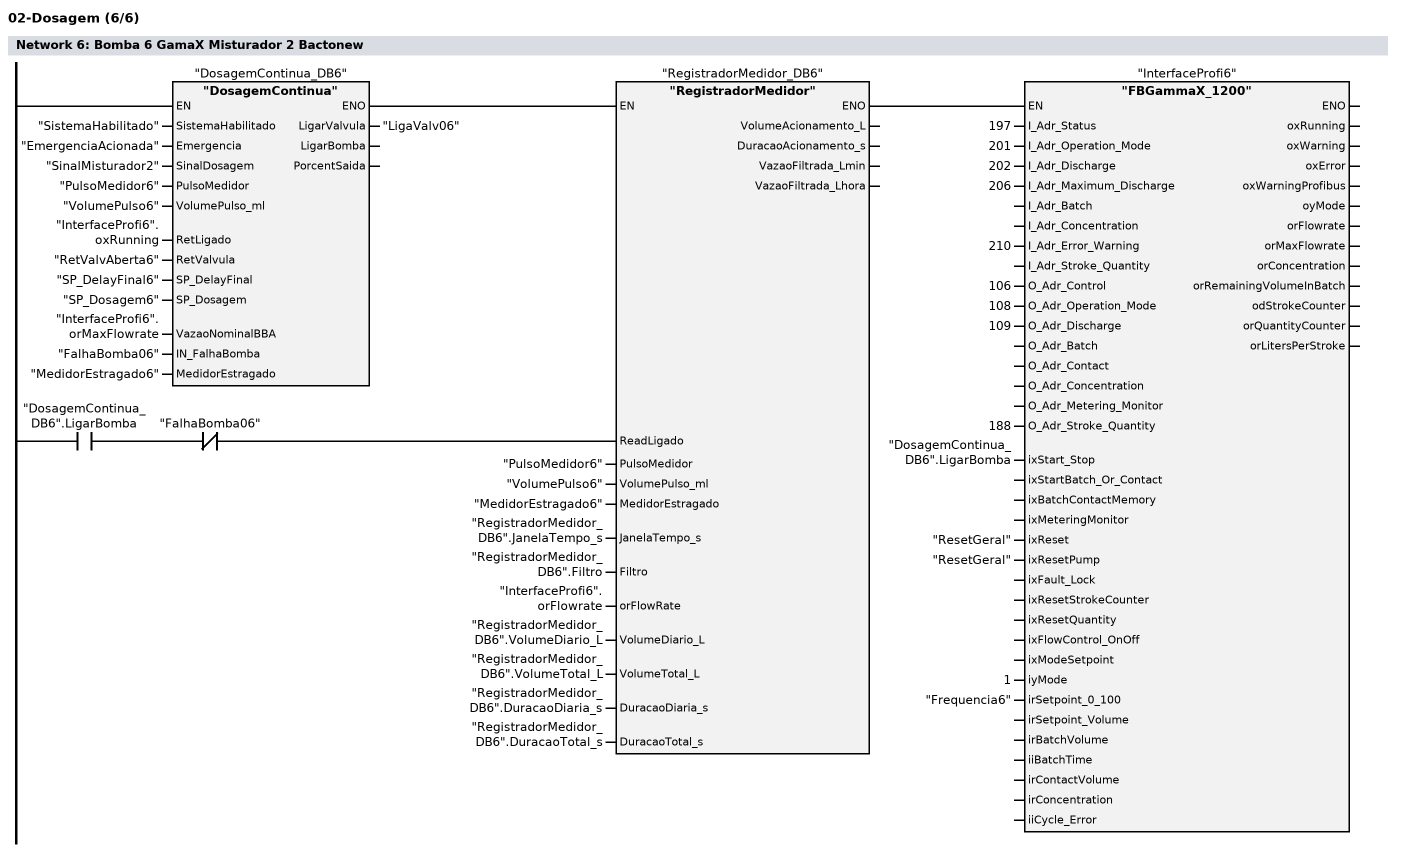
   RUNG wire#powerrail
      "DosagemContinua_DB6"(SistemaHabilitado := "SistemaHabilitado", Emergencia := "EmergenciaAcionada", SinalDosagem := "SinalMisturador2", PulsoMedidor := "PulsoMedidor6", VolumePulso_ml := "VolumePulso6", RetLigado := "InterfaceProfi6".oxRunning, RetValvula := "RetValvAberta6", SP_DelayFinal := "SP_DelayFinal6", SP_Dosagem := "SP_Dosagem6", VazaoNominalBBA := "InterfaceProfi6".orMaxFlowrate, IN_FalhaBomba := "FalhaBomba06", MedidorEstragado := "MedidorEstragado6", LigarValvula => "LigaValv06", LigarBomba =>, PorcentSaida =>)
      "RegistradorMedidor_DB6"(ReadLigado := wire#w1, PulsoMedidor := "PulsoMedidor6", VolumePulso_ml := "VolumePulso6", MedidorEstragado := "MedidorEstragado6", JanelaTempo_s := "RegistradorMedidor_DB6".JanelaTempo_s, Filtro := "RegistradorMedidor_DB6".Filtro, orFlowRate := "InterfaceProfi6".orFlowrate, VolumeDiario_L := "RegistradorMedidor_DB6".VolumeDiario_L, VolumeTotal_L := "RegistradorMedidor_DB6".VolumeTotal_L, DuracaoDiaria_s := "RegistradorMedidor_DB6".DuracaoDiaria_s, DuracaoTotal_s := "RegistradorMedidor_DB6".DuracaoTotal_s, VolumeAcionamento_L =>, DuracaoAcionamento_s =>, VazaoFiltrada_Lmin =>, VazaoFiltrada_Lhora =>)
      "InterfaceProfi6"(I_Adr_Status := 197, I_Adr_Operation_Mode := 201, I_Adr_Discharge := 202, I_Adr_Maximum_Discharge := 206, I_Adr_Batch :=, I_Adr_Concentration :=, I_Adr_Error_Warning := 210, I_Adr_Stroke_Quantity :=, O_Adr_Control := 106, O_Adr_Operation_Mode := 108, O_Adr_Discharge := 109, O_Adr_Batch :=, O_Adr_Contact :=, O_Adr_Concentration :=, O_Adr_Metering_Monitor :=, O_Adr_Stroke_Quantity := 188, ixStart_Stop := "DosagemContinua_DB6".LigarBomba, ixStartBatch_Or_Contact :=, ixBatchContactMemory :=, ixMeteringMonitor :=, ixReset := "ResetGeral", ixResetPump := "ResetGeral", ixFault_Lock :=, ixResetStrokeCounter :=, ixResetQuantity :=, ixFlowControl_OnOff :=, ixModeSetpoint :=, iyMode := 1, irSetpoint_0_100 := "Frequencia6", irSetpoint_Volume :=, irBatchVolume :=, iiBatchTime :=, irContactVolume :=, irConcentration :=, iiCycle_Error :=, oxRunning =>, oxWarning =>, oxError =>, oxWarningProfibus =>, oyMode =>, orFlowrate =>, orMaxFlowrate =>, orConcentration =>, orRemainingVolumeInBatch =>, odStrokeCounter =>, orQuantityCounter =>, orLitersPerStroke =>)
   END_RUNG
   RUNG wire#powerrail
      Contact( "DosagemContinua_DB6".LigarBomba )
      I_Contact( "FalhaBomba06" )
   END_RUNG wire#w1
   // the same network as SCL:
   "DosagemContinua_DB6"(SistemaHabilitado := "SistemaHabilitado",   // "DosagemContinua"
                         Emergencia := "EmergenciaAcionada",
                         SinalDosagem := "SinalMisturador2",
                         PulsoMedidor := "PulsoMedidor6",
                         VolumePulso_ml := "VolumePulso6",
                         RetLigado := "InterfaceProfi6".oxRunning,
                         RetValvula := "RetValvAberta6",
                         SP_DelayFinal := "SP_DelayFinal6",
                         SP_Dosagem := "SP_Dosagem6",
                         VazaoNominalBBA := "InterfaceProfi6".orMaxFlowrate,
                         IN_FalhaBomba := "FalhaBomba06",
                         MedidorEstragado := "MedidorEstragado6",
                         LigarValvula => "LigaValv06",
                         ENO => #_w1);
   "RegistradorMedidor_DB6"(EN := #_w1,   // "RegistradorMedidor"
                           ReadLigado := "DosagemContinua_DB6".LigarBomba AND NOT "FalhaBomba06",
                           PulsoMedidor := "PulsoMedidor6",
                           VolumePulso_ml := "VolumePulso6",
                           MedidorEstragado := "MedidorEstragado6",
                           JanelaTempo_s := "RegistradorMedidor_DB6".JanelaTempo_s,
                           Filtro := "RegistradorMedidor_DB6".Filtro,
                           orFlowRate := "InterfaceProfi6".orFlowrate,
                           VolumeDiario_L := "RegistradorMedidor_DB6".VolumeDiario_L,
                           VolumeTotal_L := "RegistradorMedidor_DB6".VolumeTotal_L,
                           DuracaoDiaria_s := "RegistradorMedidor_DB6".DuracaoDiaria_s,
                           DuracaoTotal_s := "RegistradorMedidor_DB6".DuracaoTotal_s,
                           ENO => #_w2);
   IF #_w2 THEN
       "InterfaceProfi6"(I_Adr_Status := 197,   // "FBGammaX_1200"
                         I_Adr_Operation_Mode := 201,
                         I_Adr_Discharge := 202,
                         I_Adr_Maximum_Discharge := 206,
                         I_Adr_Error_Warning := 210,
                         O_Adr_Control := 106,
                         O_Adr_Operation_Mode := 108,
                         O_Adr_Discharge := 109,
                         O_Adr_Stroke_Quantity := 188,
                         ixStart_Stop := "DosagemContinua_DB6".LigarBomba,
                         ixReset := "ResetGeral",
                         ixResetPump := "ResetGeral",
                         iyMode := 1,
                         irSetpoint_0_100 := "Frequencia6");
   END_IF;
END_REGION
END_ORGANIZATION_BLOCK

ORGANIZATION_BLOCK "03-Alarmes"   // OB125, LAD, ProgramCycle
TITLE = "Main Program Sweep (Cycle)"
{ S7_Optimized_Access := 'TRUE' }
VERSION : 0.1
// Alarmes e falhas de todo o sistema
   VAR_INPUT
      Initial_Call : Bool;   // Initial call of this OB
      Remanence : Bool;   // =True, if remanent data are available
   END_VAR
BEGIN

REGION Network 1: Seta falha geral
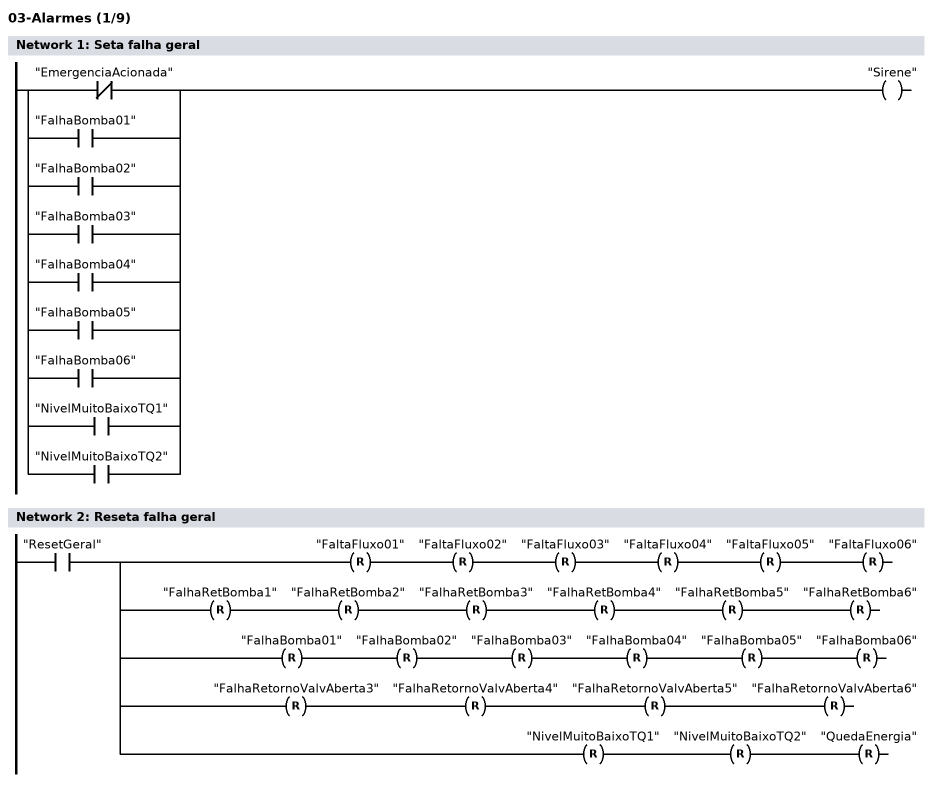
   RUNG wire#powerrail
      I_Contact( "EmergenciaAcionada" )
      wire#w1
      Coil( "Sirene" )
   END_RUNG
   RUNG wire#powerrail
      Contact( "FalhaBomba01" )
   END_RUNG wire#w1
   RUNG wire#powerrail
      Contact( "FalhaBomba02" )
   END_RUNG wire#w1
   RUNG wire#powerrail
      Contact( "FalhaBomba03" )
   END_RUNG wire#w1
   RUNG wire#powerrail
      Contact( "FalhaBomba04" )
   END_RUNG wire#w1
   RUNG wire#powerrail
      Contact( "FalhaBomba05" )
   END_RUNG wire#w1
   RUNG wire#powerrail
      Contact( "FalhaBomba06" )
   END_RUNG wire#w1
   RUNG wire#powerrail
      Contact( "NivelMuitoBaixoTQ1" )
   END_RUNG wire#w1
   RUNG wire#powerrail
      Contact( "NivelMuitoBaixoTQ2" )
   END_RUNG wire#w1
   // the same network as SCL:
   "Sirene" := NOT "EmergenciaAcionada" OR "FalhaBomba01" OR "FalhaBomba02" OR "FalhaBomba03" OR "FalhaBomba04" OR "FalhaBomba05" OR "FalhaBomba06" OR "NivelMuitoBaixoTQ1" OR "NivelMuitoBaixoTQ2";
END_REGION

REGION Network 2: Reseta falha geral
   RUNG wire#powerrail
      Contact( "ResetGeral" )
      wire#w1
      R_Coil( "FaltaFluxo01" )
      R_Coil( "FaltaFluxo02" )
      R_Coil( "FaltaFluxo03" )
      R_Coil( "FaltaFluxo04" )
      R_Coil( "FaltaFluxo05" )
      R_Coil( "FaltaFluxo06" )
   END_RUNG
   RUNG wire#w1
      R_Coil( "FalhaRetBomba1" )
      R_Coil( "FalhaRetBomba2" )
      R_Coil( "FalhaRetBomba3" )
      R_Coil( "FalhaRetBomba4" )
      R_Coil( "FalhaRetBomba5" )
      R_Coil( "FalhaRetBomba6" )
   END_RUNG
   RUNG wire#w1
      R_Coil( "FalhaBomba01" )
      R_Coil( "FalhaBomba02" )
      R_Coil( "FalhaBomba03" )
      R_Coil( "FalhaBomba04" )
      R_Coil( "FalhaBomba05" )
      R_Coil( "FalhaBomba06" )
   END_RUNG
   RUNG wire#w1
      R_Coil( "FalhaRetornoValvAberta3" )
      R_Coil( "FalhaRetornoValvAberta4" )
      R_Coil( "FalhaRetornoValvAberta5" )
      R_Coil( "FalhaRetornoValvAberta6" )
   END_RUNG
   RUNG wire#w1
      R_Coil( "NivelMuitoBaixoTQ1" )
      R_Coil( "NivelMuitoBaixoTQ2" )
      R_Coil( "QuedaEnergia" )
   END_RUNG
   // the same network as SCL:
   IF "ResetGeral" THEN
       "FaltaFluxo01" := FALSE;
       "FaltaFluxo02" := FALSE;
       "FaltaFluxo03" := FALSE;
       "FaltaFluxo04" := FALSE;
       "FaltaFluxo05" := FALSE;
       "FaltaFluxo06" := FALSE;
       "FalhaRetBomba1" := FALSE;
       "FalhaRetBomba2" := FALSE;
       "FalhaRetBomba3" := FALSE;
       "FalhaRetBomba4" := FALSE;
       "FalhaRetBomba5" := FALSE;
       "FalhaRetBomba6" := FALSE;
       "FalhaBomba01" := FALSE;
       "FalhaBomba02" := FALSE;
       "FalhaBomba03" := FALSE;
       "FalhaBomba04" := FALSE;
       "FalhaBomba05" := FALSE;
       "FalhaBomba06" := FALSE;
       "FalhaRetornoValvAberta3" := FALSE;
       "FalhaRetornoValvAberta4" := FALSE;
       "FalhaRetornoValvAberta5" := FALSE;
       "FalhaRetornoValvAberta6" := FALSE;
       "NivelMuitoBaixoTQ1" := FALSE;
       "NivelMuitoBaixoTQ2" := FALSE;
       "QuedaEnergia" := FALSE;
   END_IF;
END_REGION

REGION Network 3: Status falhas
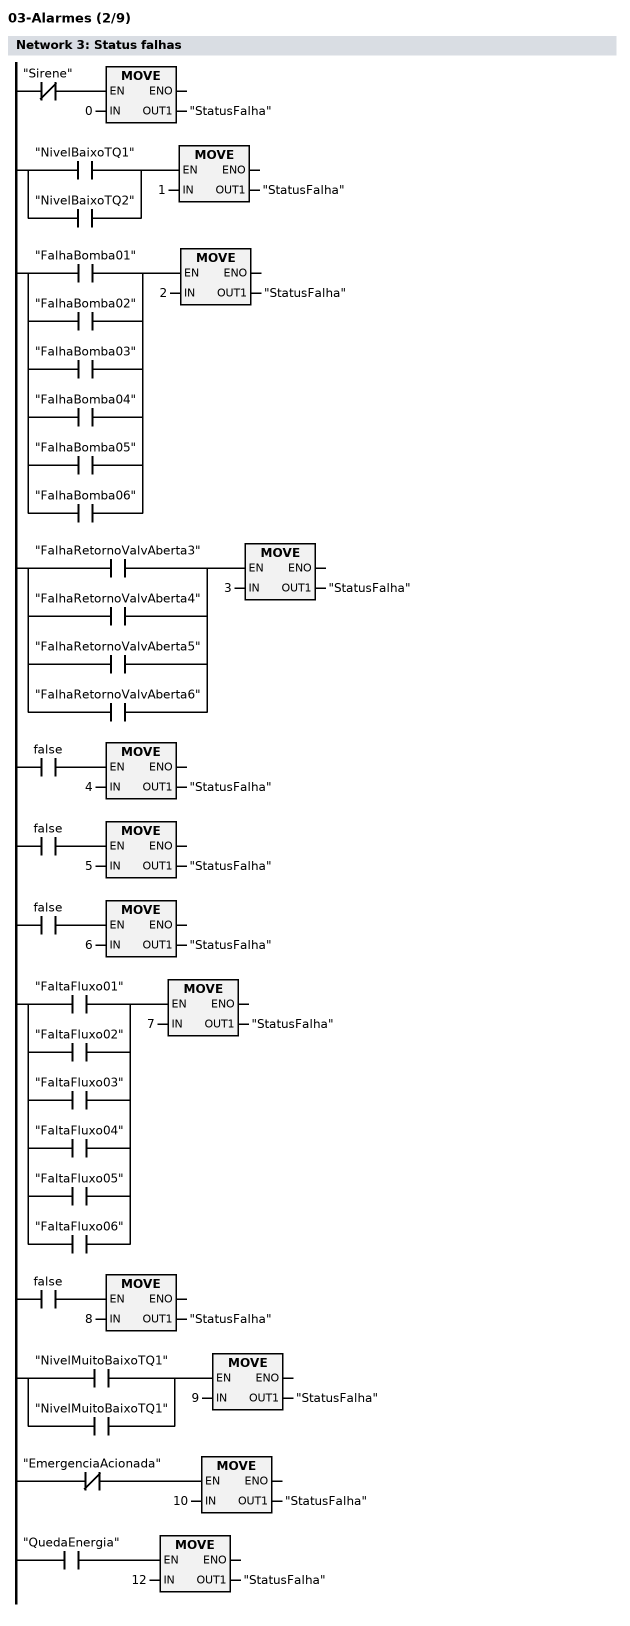
   RUNG wire#powerrail
      I_Contact( "Sirene" )
      Move(in := 0, out1 => "StatusFalha")
   END_RUNG
   RUNG wire#powerrail
      Contact( "NivelBaixoTQ1" )
      wire#w1
      Move(in := 1, out1 => "StatusFalha")
   END_RUNG
   RUNG wire#powerrail
      Contact( "NivelBaixoTQ2" )
   END_RUNG wire#w1
   RUNG wire#powerrail
      Contact( "FalhaBomba01" )
      wire#w2
      Move(in := 2, out1 => "StatusFalha")
   END_RUNG
   RUNG wire#powerrail
      Contact( "FalhaBomba02" )
   END_RUNG wire#w2
   RUNG wire#powerrail
      Contact( "FalhaBomba03" )
   END_RUNG wire#w2
   RUNG wire#powerrail
      Contact( "FalhaBomba04" )
   END_RUNG wire#w2
   RUNG wire#powerrail
      Contact( "FalhaBomba05" )
   END_RUNG wire#w2
   RUNG wire#powerrail
      Contact( "FalhaBomba06" )
   END_RUNG wire#w2
   RUNG wire#powerrail
      Contact( "FalhaRetornoValvAberta3" )
      wire#w3
      Move(in := 3, out1 => "StatusFalha")
   END_RUNG
   RUNG wire#powerrail
      Contact( "FalhaRetornoValvAberta4" )
   END_RUNG wire#w3
   RUNG wire#powerrail
      Contact( "FalhaRetornoValvAberta5" )
   END_RUNG wire#w3
   RUNG wire#powerrail
      Contact( "FalhaRetornoValvAberta6" )
   END_RUNG wire#w3
   RUNG wire#powerrail
      Contact( false )
      Move(in := 4, out1 => "StatusFalha")
   END_RUNG
   RUNG wire#powerrail
      Contact( false )
      Move(in := 5, out1 => "StatusFalha")
   END_RUNG
   RUNG wire#powerrail
      Contact( false )
      Move(in := 6, out1 => "StatusFalha")
   END_RUNG
   RUNG wire#powerrail
      Contact( "FaltaFluxo01" )
      wire#w4
      Move(in := 7, out1 => "StatusFalha")
   END_RUNG
   RUNG wire#powerrail
      Contact( "FaltaFluxo02" )
   END_RUNG wire#w4
   RUNG wire#powerrail
      Contact( "FaltaFluxo03" )
   END_RUNG wire#w4
   RUNG wire#powerrail
      Contact( "FaltaFluxo04" )
   END_RUNG wire#w4
   RUNG wire#powerrail
      Contact( "FaltaFluxo05" )
   END_RUNG wire#w4
   RUNG wire#powerrail
      Contact( "FaltaFluxo06" )
   END_RUNG wire#w4
   RUNG wire#powerrail
      Contact( false )
      Move(in := 8, out1 => "StatusFalha")
   END_RUNG
   RUNG wire#powerrail
      Contact( "NivelMuitoBaixoTQ1" )
      wire#w5
      Move(in := 9, out1 => "StatusFalha")
   END_RUNG
   RUNG wire#powerrail
      Contact( "NivelMuitoBaixoTQ1" )
   END_RUNG wire#w5
   RUNG wire#powerrail
      I_Contact( "EmergenciaAcionada" )
      Move(in := 10, out1 => "StatusFalha")
   END_RUNG
   RUNG wire#powerrail
      Contact( "QuedaEnergia" )
      Move(in := 12, out1 => "StatusFalha")
   END_RUNG
   // the same network as SCL:
   IF NOT "Sirene" THEN "StatusFalha" := 0; END_IF;
   IF "NivelBaixoTQ1" OR "NivelBaixoTQ2" THEN "StatusFalha" := 1; END_IF;
   IF "FalhaBomba01" OR "FalhaBomba02" OR "FalhaBomba03" OR "FalhaBomba04" OR "FalhaBomba05" OR "FalhaBomba06" THEN
       "StatusFalha" := 2;
   END_IF;
   IF "FalhaRetornoValvAberta3" OR "FalhaRetornoValvAberta4" OR "FalhaRetornoValvAberta5" OR "FalhaRetornoValvAberta6" THEN
       "StatusFalha" := 3;
   END_IF;
   IF false THEN
       "StatusFalha" := 4;
       "StatusFalha" := 5;
       "StatusFalha" := 6;
   END_IF;
   IF "FaltaFluxo01" OR "FaltaFluxo02" OR "FaltaFluxo03" OR "FaltaFluxo04" OR "FaltaFluxo05" OR "FaltaFluxo06" THEN
       "StatusFalha" := 7;
   END_IF;
   IF false THEN "StatusFalha" := 8; END_IF;
   IF "NivelMuitoBaixoTQ1" OR "NivelMuitoBaixoTQ1" THEN "StatusFalha" := 9; END_IF;
   IF NOT "EmergenciaAcionada" THEN "StatusFalha" := 10; END_IF;
   IF "QuedaEnergia" THEN "StatusFalha" := 12; END_IF;
END_REGION

REGION Network 4: Falhas Bomba 01
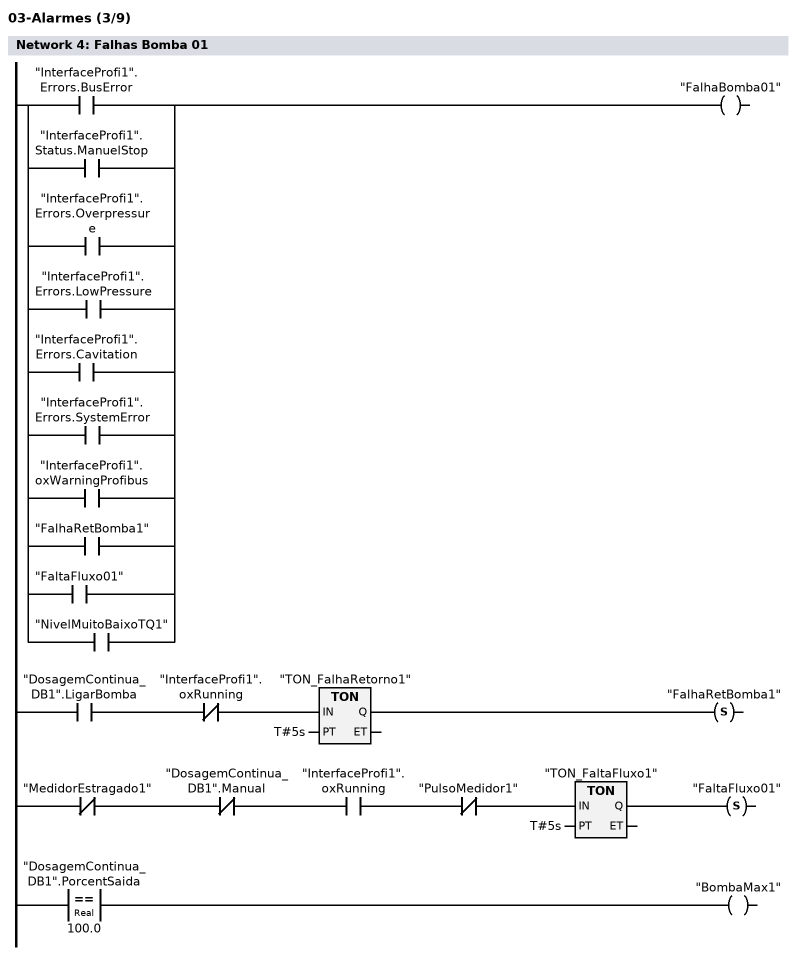
   "FalhaBomba01" := "InterfaceProfi1".Errors.BusError OR "InterfaceProfi1".Status.ManuelStop OR "InterfaceProfi1".Errors.Overpressure OR "InterfaceProfi1".Errors.LowPressure OR "InterfaceProfi1".Errors.Cavitation OR "InterfaceProfi1".Errors.SystemError OR "InterfaceProfi1".oxWarningProfibus OR "FalhaRetBomba1" OR "FaltaFluxo01" OR "NivelMuitoBaixoTQ1";
   "TON_FalhaRetorno1".TON(IN := "DosagemContinua_DB1".LigarBomba AND NOT "InterfaceProfi1".oxRunning,
                           PT := T#5s);
   IF "TON_FalhaRetorno1".Q THEN "FalhaRetBomba1" := TRUE; END_IF;
   "TON_FaltaFluxo1".TON(IN := NOT "MedidorEstragado1" AND NOT "DosagemContinua_DB1".Manual AND "InterfaceProfi1".oxRunning AND NOT "PulsoMedidor1",
                         PT := T#5s);
   IF "TON_FaltaFluxo1".Q THEN "FaltaFluxo01" := TRUE; END_IF;
   "BombaMax1" := "DosagemContinua_DB1".PorcentSaida = 100.0;
END_REGION

REGION Network 5: Falhas Bomba 02
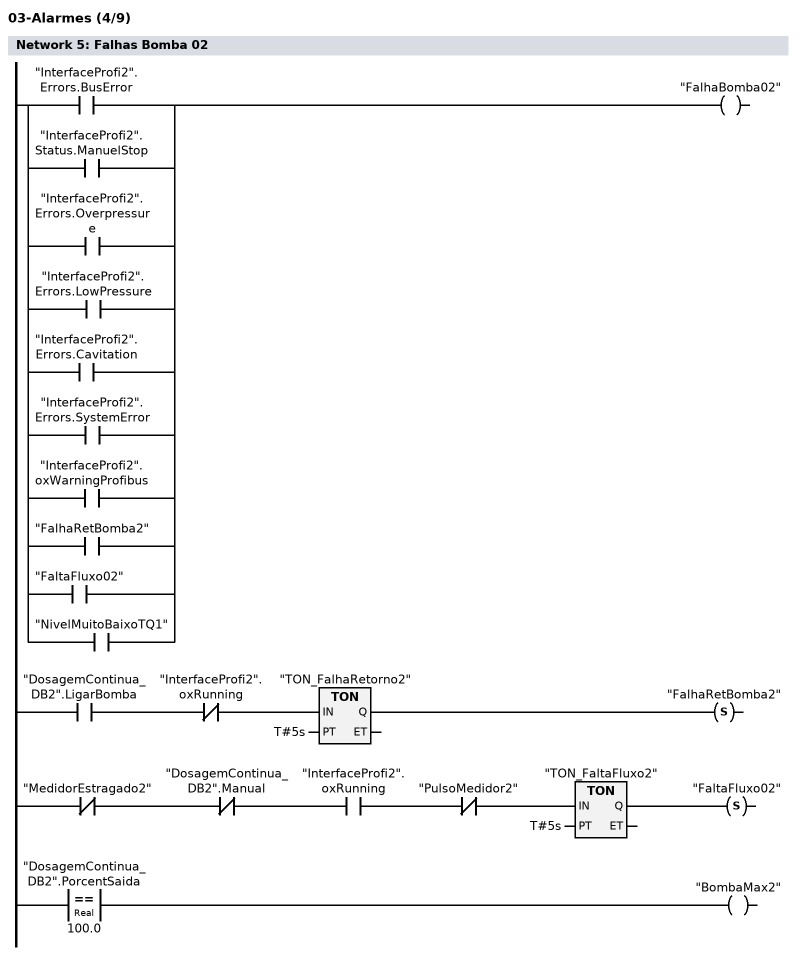
   "FalhaBomba02" := "InterfaceProfi2".Errors.BusError OR "InterfaceProfi2".Status.ManuelStop OR "InterfaceProfi2".Errors.Overpressure OR "InterfaceProfi2".Errors.LowPressure OR "InterfaceProfi2".Errors.Cavitation OR "InterfaceProfi2".Errors.SystemError OR "InterfaceProfi2".oxWarningProfibus OR "FalhaRetBomba2" OR "FaltaFluxo02" OR "NivelMuitoBaixoTQ1";
   "TON_FalhaRetorno2".TON(IN := "DosagemContinua_DB2".LigarBomba AND NOT "InterfaceProfi2".oxRunning,
                           PT := T#5s);
   IF "TON_FalhaRetorno2".Q THEN "FalhaRetBomba2" := TRUE; END_IF;
   "TON_FaltaFluxo2".TON(IN := NOT "MedidorEstragado2" AND NOT "DosagemContinua_DB2".Manual AND "InterfaceProfi2".oxRunning AND NOT "PulsoMedidor2",
                         PT := T#5s);
   IF "TON_FaltaFluxo2".Q THEN "FaltaFluxo02" := TRUE; END_IF;
   "BombaMax2" := "DosagemContinua_DB2".PorcentSaida = 100.0;
END_REGION

REGION Network 6: Falhas Bomba 03
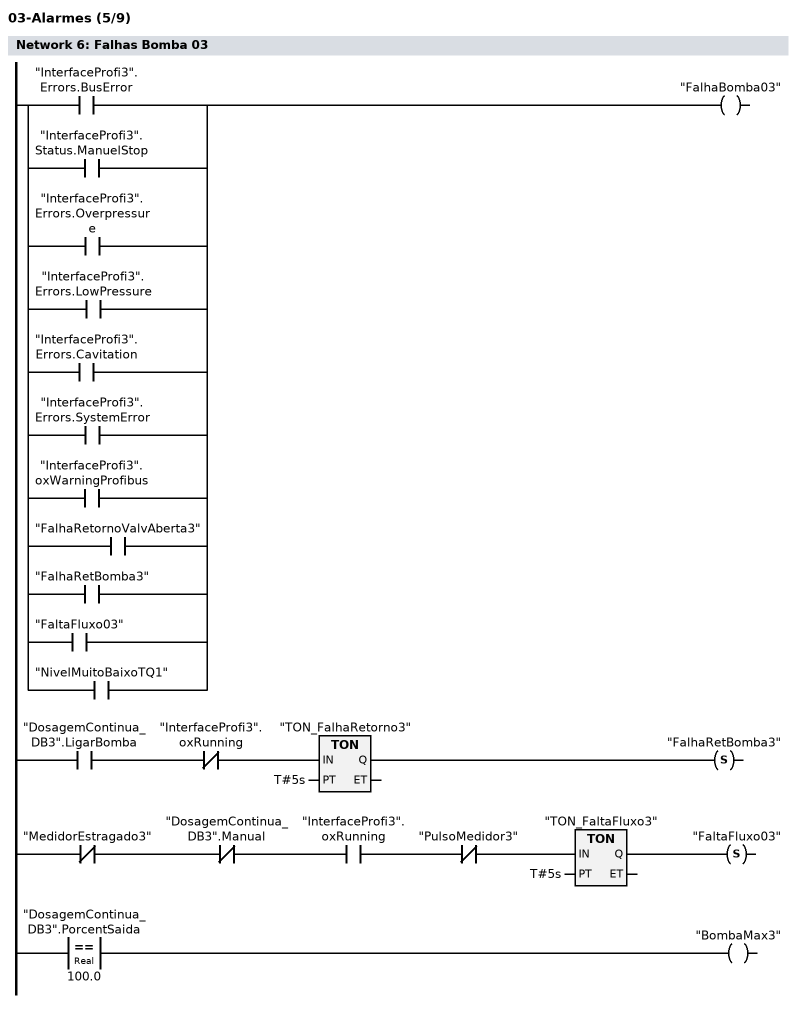
   "FalhaBomba03" := "InterfaceProfi3".Errors.BusError OR "InterfaceProfi3".Status.ManuelStop OR "InterfaceProfi3".Errors.Overpressure OR "InterfaceProfi3".Errors.LowPressure OR "InterfaceProfi3".Errors.Cavitation OR "InterfaceProfi3".Errors.SystemError OR "InterfaceProfi3".oxWarningProfibus OR "FalhaRetornoValvAberta3" OR "FalhaRetBomba3" OR "FaltaFluxo03" OR "NivelMuitoBaixoTQ1";
   "TON_FalhaRetorno3".TON(IN := "DosagemContinua_DB3".LigarBomba AND NOT "InterfaceProfi3".oxRunning,
                           PT := T#5s);
   IF "TON_FalhaRetorno3".Q THEN "FalhaRetBomba3" := TRUE; END_IF;
   "TON_FaltaFluxo3".TON(IN := NOT "MedidorEstragado3" AND NOT "DosagemContinua_DB3".Manual AND "InterfaceProfi3".oxRunning AND NOT "PulsoMedidor3",
                         PT := T#5s);
   IF "TON_FaltaFluxo3".Q THEN "FaltaFluxo03" := TRUE; END_IF;
   "BombaMax3" := "DosagemContinua_DB3".PorcentSaida = 100.0;
END_REGION

REGION Network 7: Falhas Bomba 04
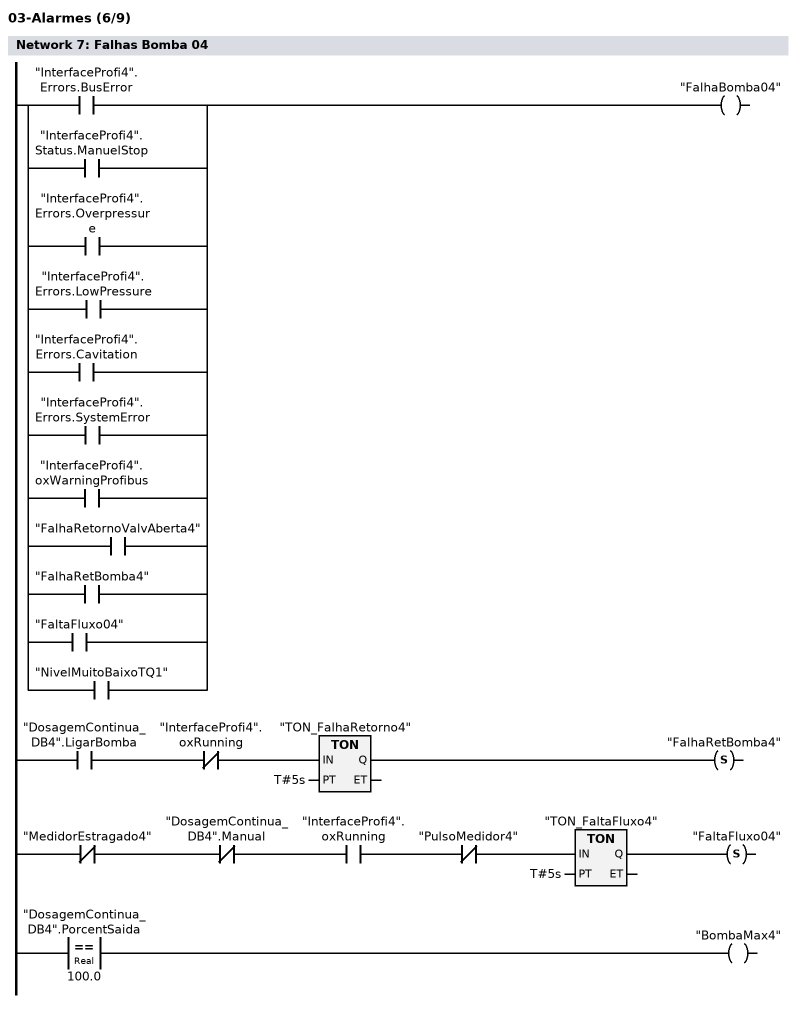
   "FalhaBomba04" := "InterfaceProfi4".Errors.BusError OR "InterfaceProfi4".Status.ManuelStop OR "InterfaceProfi4".Errors.Overpressure OR "InterfaceProfi4".Errors.LowPressure OR "InterfaceProfi4".Errors.Cavitation OR "InterfaceProfi4".Errors.SystemError OR "InterfaceProfi4".oxWarningProfibus OR "FalhaRetornoValvAberta4" OR "FalhaRetBomba4" OR "FaltaFluxo04" OR "NivelMuitoBaixoTQ1";
   "TON_FalhaRetorno4".TON(IN := "DosagemContinua_DB4".LigarBomba AND NOT "InterfaceProfi4".oxRunning,
                           PT := T#5s);
   IF "TON_FalhaRetorno4".Q THEN "FalhaRetBomba4" := TRUE; END_IF;
   "TON_FaltaFluxo4".TON(IN := NOT "MedidorEstragado4" AND NOT "DosagemContinua_DB4".Manual AND "InterfaceProfi4".oxRunning AND NOT "PulsoMedidor4",
                         PT := T#5s);
   IF "TON_FaltaFluxo4".Q THEN "FaltaFluxo04" := TRUE; END_IF;
   "BombaMax4" := "DosagemContinua_DB4".PorcentSaida = 100.0;
END_REGION

REGION Network 8: Falhas Bomba 05
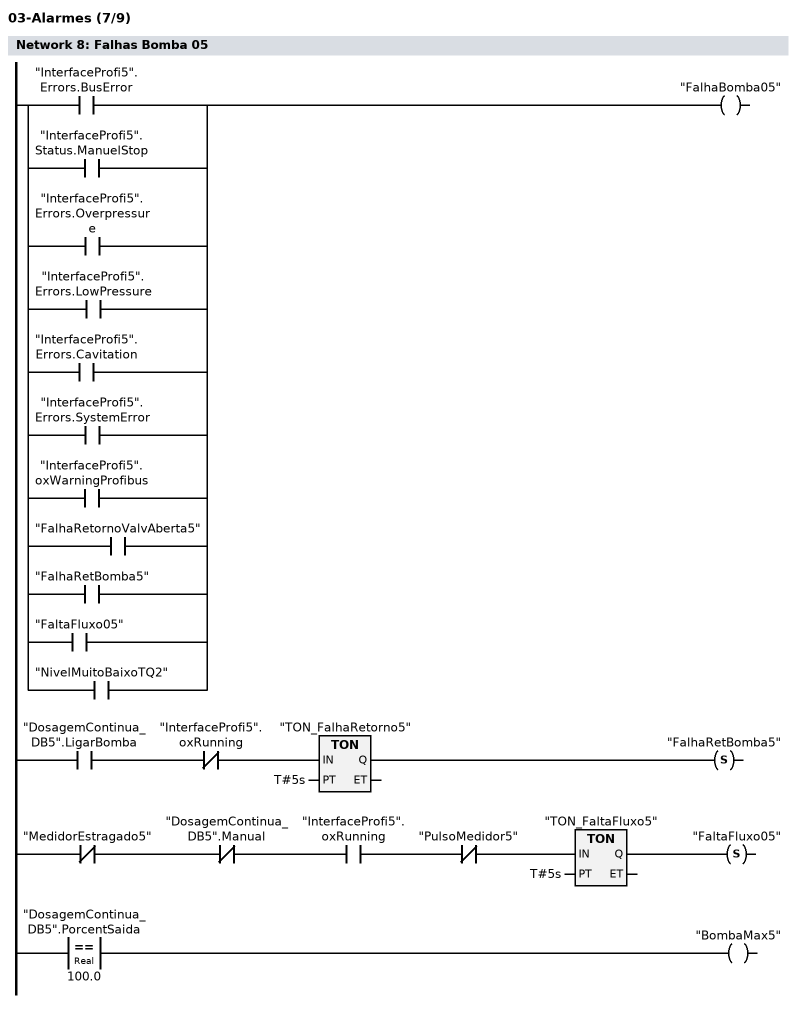
   "FalhaBomba05" := "InterfaceProfi5".Errors.BusError OR "InterfaceProfi5".Status.ManuelStop OR "InterfaceProfi5".Errors.Overpressure OR "InterfaceProfi5".Errors.LowPressure OR "InterfaceProfi5".Errors.Cavitation OR "InterfaceProfi5".Errors.SystemError OR "InterfaceProfi5".oxWarningProfibus OR "FalhaRetornoValvAberta5" OR "FalhaRetBomba5" OR "FaltaFluxo05" OR "NivelMuitoBaixoTQ2";
   "TON_FalhaRetorno5".TON(IN := "DosagemContinua_DB5".LigarBomba AND NOT "InterfaceProfi5".oxRunning,
                           PT := T#5s);
   IF "TON_FalhaRetorno5".Q THEN "FalhaRetBomba5" := TRUE; END_IF;
   "TON_FaltaFluxo5".TON(IN := NOT "MedidorEstragado5" AND NOT "DosagemContinua_DB5".Manual AND "InterfaceProfi5".oxRunning AND NOT "PulsoMedidor5",
                         PT := T#5s);
   IF "TON_FaltaFluxo5".Q THEN "FaltaFluxo05" := TRUE; END_IF;
   "BombaMax5" := "DosagemContinua_DB5".PorcentSaida = 100.0;
END_REGION

REGION Network 9: Falhas Bomba 06
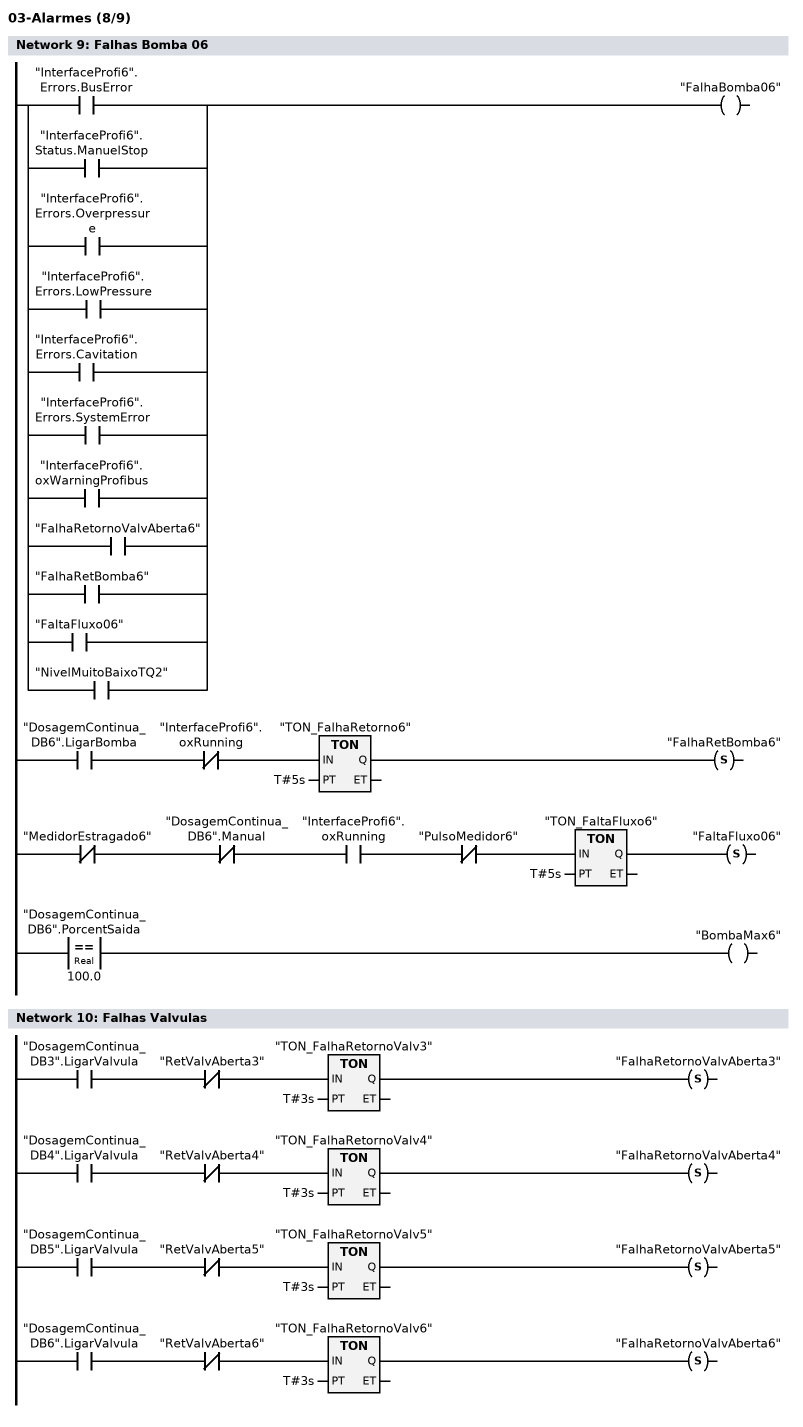
   "FalhaBomba06" := "InterfaceProfi6".Errors.BusError OR "InterfaceProfi6".Status.ManuelStop OR "InterfaceProfi6".Errors.Overpressure OR "InterfaceProfi6".Errors.LowPressure OR "InterfaceProfi6".Errors.Cavitation OR "InterfaceProfi6".Errors.SystemError OR "InterfaceProfi6".oxWarningProfibus OR "FalhaRetornoValvAberta6" OR "FalhaRetBomba6" OR "FaltaFluxo06" OR "NivelMuitoBaixoTQ2";
   "TON_FalhaRetorno6".TON(IN := "DosagemContinua_DB6".LigarBomba AND NOT "InterfaceProfi6".oxRunning,
                           PT := T#5s);
   IF "TON_FalhaRetorno6".Q THEN "FalhaRetBomba6" := TRUE; END_IF;
   "TON_FaltaFluxo6".TON(IN := NOT "MedidorEstragado6" AND NOT "DosagemContinua_DB6".Manual AND "InterfaceProfi6".oxRunning AND NOT "PulsoMedidor6",
                         PT := T#5s);
   IF "TON_FaltaFluxo6".Q THEN "FaltaFluxo06" := TRUE; END_IF;
   "BombaMax6" := "DosagemContinua_DB6".PorcentSaida = 100.0;
END_REGION

REGION Network 10: Falhas Valvulas
   "TON_FalhaRetornoValv3".TON(IN := "DosagemContinua_DB3".LigarValvula AND NOT "RetValvAberta3", PT := T#3s);
   IF "TON_FalhaRetornoValv3".Q THEN "FalhaRetornoValvAberta3" := TRUE; END_IF;
   "TON_FalhaRetornoValv4".TON(IN := "DosagemContinua_DB4".LigarValvula AND NOT "RetValvAberta4", PT := T#3s);
   IF "TON_FalhaRetornoValv4".Q THEN "FalhaRetornoValvAberta4" := TRUE; END_IF;
   "TON_FalhaRetornoValv5".TON(IN := "DosagemContinua_DB5".LigarValvula AND NOT "RetValvAberta5", PT := T#3s);
   IF "TON_FalhaRetornoValv5".Q THEN "FalhaRetornoValvAberta5" := TRUE; END_IF;
   "TON_FalhaRetornoValv6".TON(IN := "DosagemContinua_DB6".LigarValvula AND NOT "RetValvAberta6", PT := T#3s);
   IF "TON_FalhaRetornoValv6".Q THEN "FalhaRetornoValvAberta6" := TRUE; END_IF;
END_REGION

REGION Network 11: Nivel baixo dos tanques
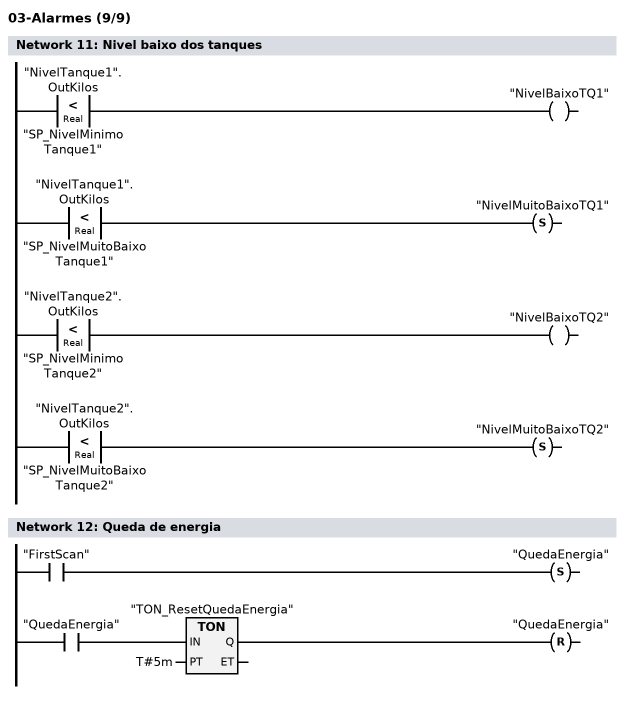
   RUNG wire#powerrail
      { S7_Templates := "SrcType := Real" } LT_Contact(in1 := "NivelTanque1".OutKilos, in2 := "SP_NivelMinimoTanque1")
      Coil( "NivelBaixoTQ1" )
   END_RUNG
   RUNG wire#powerrail
      { S7_Templates := "SrcType := Real" } LT_Contact(in1 := "NivelTanque1".OutKilos, in2 := "SP_NivelMuitoBaixoTanque1")
      S_Coil( "NivelMuitoBaixoTQ1" )
   END_RUNG
   RUNG wire#powerrail
      { S7_Templates := "SrcType := Real" } LT_Contact(in1 := "NivelTanque2".OutKilos, in2 := "SP_NivelMinimoTanque2")
      Coil( "NivelBaixoTQ2" )
   END_RUNG
   RUNG wire#powerrail
      { S7_Templates := "SrcType := Real" } LT_Contact(in1 := "NivelTanque2".OutKilos, in2 := "SP_NivelMuitoBaixoTanque2")
      S_Coil( "NivelMuitoBaixoTQ2" )
   END_RUNG
   // the same network as SCL:
   "NivelBaixoTQ1" := "NivelTanque1".OutKilos < "SP_NivelMinimoTanque1";
   IF "NivelTanque1".OutKilos < "SP_NivelMuitoBaixoTanque1" THEN "NivelMuitoBaixoTQ1" := TRUE; END_IF;
   "NivelBaixoTQ2" := "NivelTanque2".OutKilos < "SP_NivelMinimoTanque2";
   IF "NivelTanque2".OutKilos < "SP_NivelMuitoBaixoTanque2" THEN "NivelMuitoBaixoTQ2" := TRUE; END_IF;
END_REGION

REGION Network 12: Queda de energia
   IF "FirstScan" THEN "QuedaEnergia" := TRUE; END_IF;
   "TON_ResetQuedaEnergia".TON(IN := "QuedaEnergia", PT := T#5m);
   IF "TON_ResetQuedaEnergia".Q THEN "QuedaEnergia" := FALSE; END_IF;
END_REGION
END_ORGANIZATION_BLOCK

ORGANIZATION_BLOCK "04-Relatorios"   // OB126, LAD, ProgramCycle
TITLE = "Main Program Sweep (Cycle)"
{ S7_Optimized_Access := 'TRUE' }
VERSION : 0.1
   VAR_INPUT
      Initial_Call : Bool;   // Initial call of this OB
      Remanence : Bool;   // =True, if remanent data are available
   END_VAR
   VAR_TEMP   // added for the SCL form of the ladder/FBD networks
      _w1 : Bool;
      _w2 : Bool;
      _w3 : Bool;
      _w4 : Bool;
      _w5 : Bool;
      _w6 : Bool;
   END_VAR
BEGIN

REGION Network 1: Data e Hora do CLP
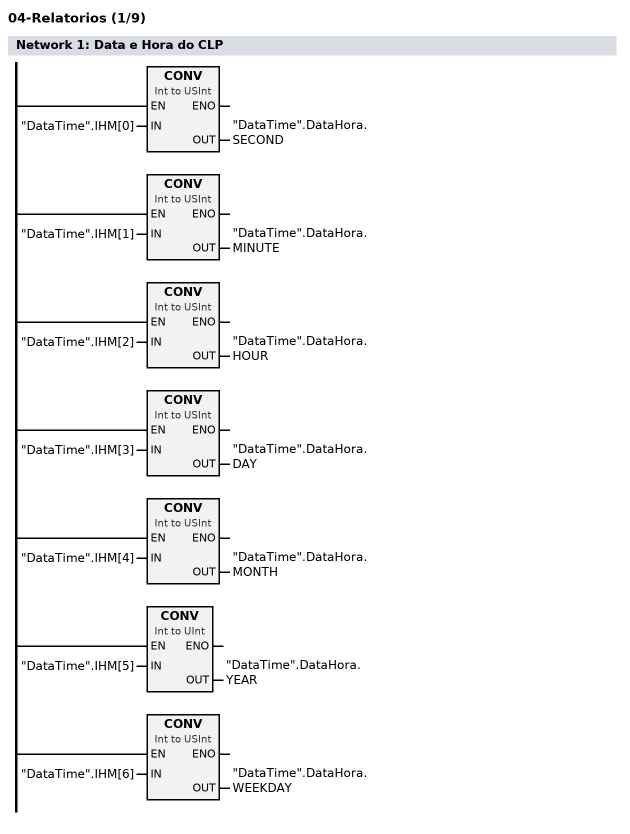
   RUNG wire#powerrail
      { S7_Templates := "[SrcType := Int, DestType := USInt]" } Convert(in := "DataTime".IHM[0], out => "DataTime".DataHora.SECOND)
   END_RUNG
   RUNG wire#powerrail
      { S7_Templates := "[SrcType := Int, DestType := USInt]" } Convert(in := "DataTime".IHM[1], out => "DataTime".DataHora.MINUTE)
   END_RUNG
   RUNG wire#powerrail
      { S7_Templates := "[SrcType := Int, DestType := USInt]" } Convert(in := "DataTime".IHM[2], out => "DataTime".DataHora.HOUR)
   END_RUNG
   RUNG wire#powerrail
      { S7_Templates := "[SrcType := Int, DestType := USInt]" } Convert(in := "DataTime".IHM[3], out => "DataTime".DataHora.DAY)
   END_RUNG
   RUNG wire#powerrail
      { S7_Templates := "[SrcType := Int, DestType := USInt]" } Convert(in := "DataTime".IHM[4], out => "DataTime".DataHora.MONTH)
   END_RUNG
   RUNG wire#powerrail
      { S7_Templates := "[SrcType := Int, DestType := UInt]" } Convert(in := "DataTime".IHM[5], out => "DataTime".DataHora.YEAR)
   END_RUNG
   RUNG wire#powerrail
      { S7_Templates := "[SrcType := Int, DestType := USInt]" } Convert(in := "DataTime".IHM[6], out => "DataTime".DataHora.WEEKDAY)
   END_RUNG
   // the same network as SCL:
   "DataTime".DataHora.SECOND := INT_TO_USINT("DataTime".IHM[0]);
   "DataTime".DataHora.MINUTE := INT_TO_USINT("DataTime".IHM[1]);
   "DataTime".DataHora.HOUR := INT_TO_USINT("DataTime".IHM[2]);
   "DataTime".DataHora.DAY := INT_TO_USINT("DataTime".IHM[3]);
   "DataTime".DataHora.MONTH := INT_TO_USINT("DataTime".IHM[4]);
   "DataTime".DataHora.YEAR := INT_TO_UINT("DataTime".IHM[5]);
   "DataTime".DataHora.WEEKDAY := INT_TO_USINT("DataTime".IHM[6]);
END_REGION

REGION Network 2: Relatorio Diario Unificado
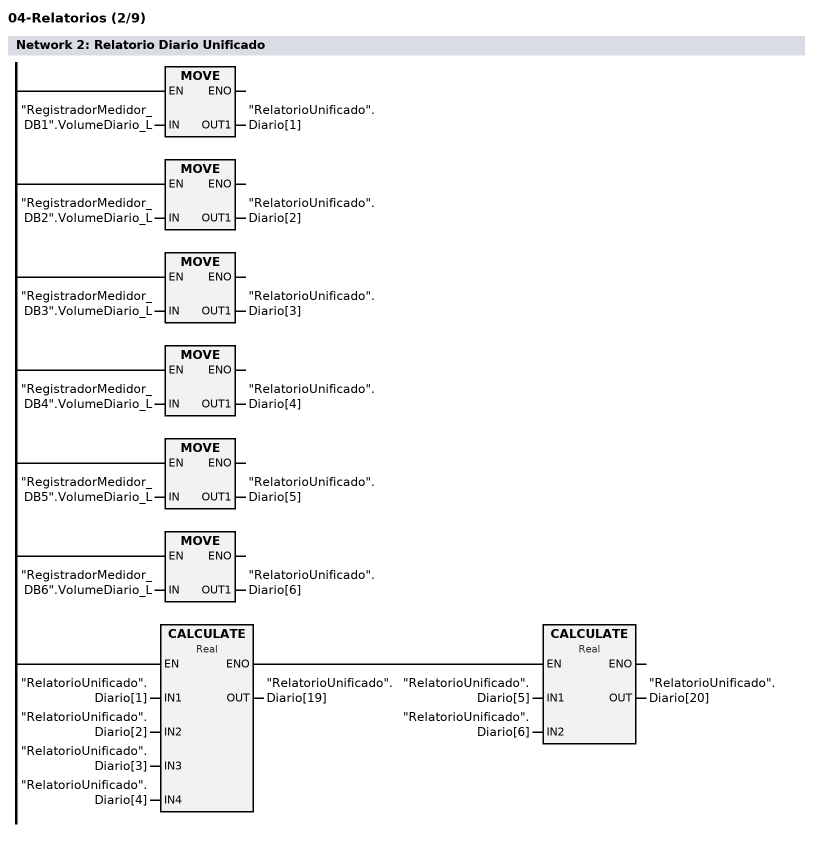
   RUNG wire#powerrail
      Move(in := "RegistradorMedidor_DB1".VolumeDiario_L, out1 => "RelatorioUnificado".Diario[1])
   END_RUNG
   RUNG wire#powerrail
      Move(in := "RegistradorMedidor_DB2".VolumeDiario_L, out1 => "RelatorioUnificado".Diario[2])
   END_RUNG
   RUNG wire#powerrail
      Move(in := "RegistradorMedidor_DB3".VolumeDiario_L, out1 => "RelatorioUnificado".Diario[3])
   END_RUNG
   RUNG wire#powerrail
      Move(in := "RegistradorMedidor_DB4".VolumeDiario_L, out1 => "RelatorioUnificado".Diario[4])
   END_RUNG
   RUNG wire#powerrail
      Move(in := "RegistradorMedidor_DB5".VolumeDiario_L, out1 => "RelatorioUnificado".Diario[5])
   END_RUNG
   RUNG wire#powerrail
      Move(in := "RegistradorMedidor_DB6".VolumeDiario_L, out1 => "RelatorioUnificado".Diario[6])
   END_RUNG
   RUNG wire#powerrail
      { S7_Templates := "SrcType := Real"; S7_Expression := "IN1 + IN2 + IN3 + IN4" } Calculate(in1 := "RelatorioUnificado".Diario[1], in2 := "RelatorioUnificado".Diario[2], in3 := "RelatorioUnificado".Diario[3], in4 := "RelatorioUnificado".Diario[4], out => "RelatorioUnificado".Diario[19])
      { S7_Templates := "SrcType := Real"; S7_Expression := "IN1 + IN2" } Calculate(in1 := "RelatorioUnificado".Diario[5], in2 := "RelatorioUnificado".Diario[6], out => "RelatorioUnificado".Diario[20])
   END_RUNG
   // the same network as SCL:
   "RelatorioUnificado".Diario[1] := "RegistradorMedidor_DB1".VolumeDiario_L;
   "RelatorioUnificado".Diario[2] := "RegistradorMedidor_DB2".VolumeDiario_L;
   "RelatorioUnificado".Diario[3] := "RegistradorMedidor_DB3".VolumeDiario_L;
   "RelatorioUnificado".Diario[4] := "RegistradorMedidor_DB4".VolumeDiario_L;
   "RelatorioUnificado".Diario[5] := "RegistradorMedidor_DB5".VolumeDiario_L;
   "RelatorioUnificado".Diario[6] := "RegistradorMedidor_DB6".VolumeDiario_L;
   "RelatorioUnificado".Diario[19] := "RelatorioUnificado".Diario[1] + "RelatorioUnificado".Diario[2] + "RelatorioUnificado".Diario[3] + "RelatorioUnificado".Diario[4];
   "RelatorioUnificado".Diario[20] := "RelatorioUnificado".Diario[5] + "RelatorioUnificado".Diario[6];
END_REGION

REGION Network 3: Vazão atual / SP Atual
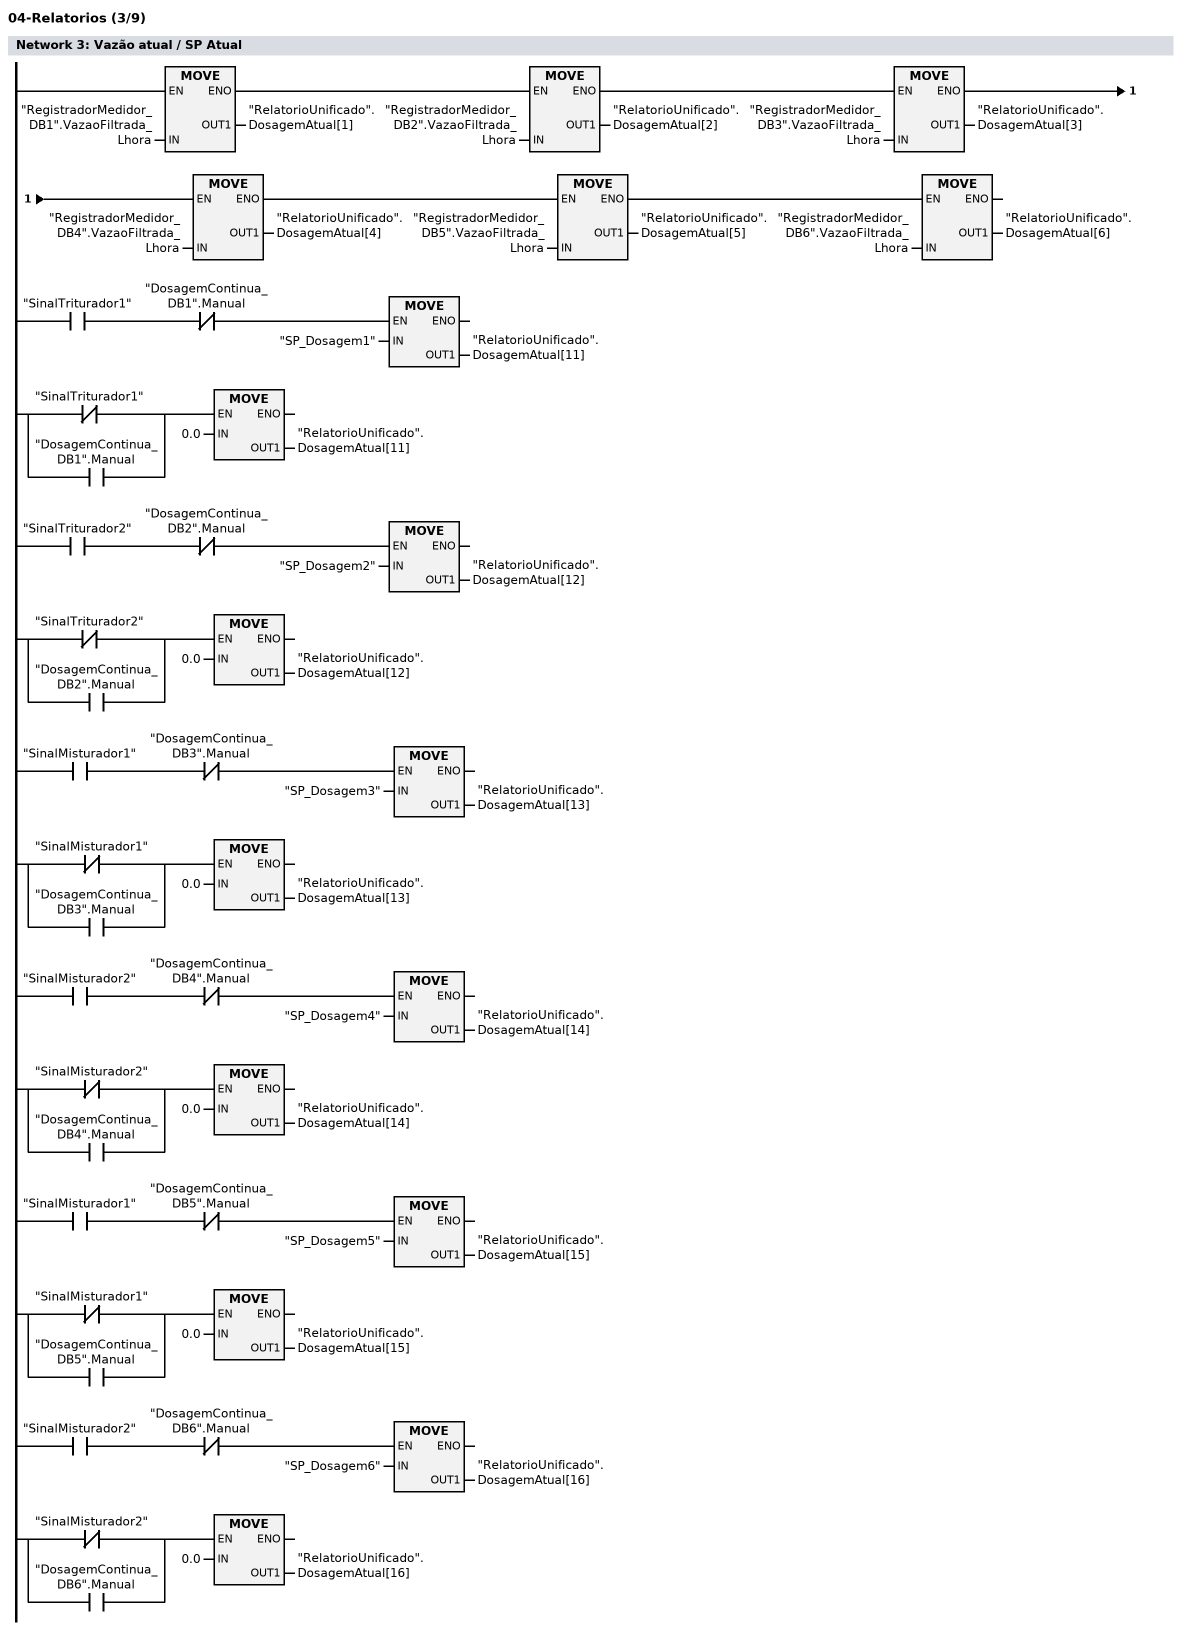
   RUNG wire#powerrail
      Move(in := "RegistradorMedidor_DB1".VazaoFiltrada_Lhora, out1 => "RelatorioUnificado".DosagemAtual[1])
      Move(in := "RegistradorMedidor_DB2".VazaoFiltrada_Lhora, out1 => "RelatorioUnificado".DosagemAtual[2])
      Move(in := "RegistradorMedidor_DB3".VazaoFiltrada_Lhora, out1 => "RelatorioUnificado".DosagemAtual[3])
      Move(in := "RegistradorMedidor_DB4".VazaoFiltrada_Lhora, out1 => "RelatorioUnificado".DosagemAtual[4])
      Move(in := "RegistradorMedidor_DB5".VazaoFiltrada_Lhora, out1 => "RelatorioUnificado".DosagemAtual[5])
      Move(in := "RegistradorMedidor_DB6".VazaoFiltrada_Lhora, out1 => "RelatorioUnificado".DosagemAtual[6])
   END_RUNG
   RUNG wire#powerrail
      Contact( "SinalTriturador1" )
      I_Contact( "DosagemContinua_DB1".Manual )
      Move(in := "SP_Dosagem1", out1 => "RelatorioUnificado".DosagemAtual[11])
   END_RUNG
   RUNG wire#powerrail
      I_Contact( "SinalTriturador1" )
      wire#w1
      Move(in := 0.0, out1 => "RelatorioUnificado".DosagemAtual[11])
   END_RUNG
   RUNG wire#powerrail
      Contact( "DosagemContinua_DB1".Manual )
   END_RUNG wire#w1
   RUNG wire#powerrail
      Contact( "SinalTriturador2" )
      I_Contact( "DosagemContinua_DB2".Manual )
      Move(in := "SP_Dosagem2", out1 => "RelatorioUnificado".DosagemAtual[12])
   END_RUNG
   RUNG wire#powerrail
      I_Contact( "SinalTriturador2" )
      wire#w2
      Move(in := 0.0, out1 => "RelatorioUnificado".DosagemAtual[12])
   END_RUNG
   RUNG wire#powerrail
      Contact( "DosagemContinua_DB2".Manual )
   END_RUNG wire#w2
   RUNG wire#powerrail
      Contact( "SinalMisturador1" )
      I_Contact( "DosagemContinua_DB3".Manual )
      Move(in := "SP_Dosagem3", out1 => "RelatorioUnificado".DosagemAtual[13])
   END_RUNG
   RUNG wire#powerrail
      I_Contact( "SinalMisturador1" )
      wire#w3
      Move(in := 0.0, out1 => "RelatorioUnificado".DosagemAtual[13])
   END_RUNG
   RUNG wire#powerrail
      Contact( "DosagemContinua_DB3".Manual )
   END_RUNG wire#w3
   RUNG wire#powerrail
      Contact( "SinalMisturador2" )
      I_Contact( "DosagemContinua_DB4".Manual )
      Move(in := "SP_Dosagem4", out1 => "RelatorioUnificado".DosagemAtual[14])
   END_RUNG
   RUNG wire#powerrail
      I_Contact( "SinalMisturador2" )
      wire#w4
      Move(in := 0.0, out1 => "RelatorioUnificado".DosagemAtual[14])
   END_RUNG
   RUNG wire#powerrail
      Contact( "DosagemContinua_DB4".Manual )
   END_RUNG wire#w4
   RUNG wire#powerrail
      Contact( "SinalMisturador1" )
      I_Contact( "DosagemContinua_DB5".Manual )
      Move(in := "SP_Dosagem5", out1 => "RelatorioUnificado".DosagemAtual[15])
   END_RUNG
   RUNG wire#powerrail
      I_Contact( "SinalMisturador1" )
      wire#w5
      Move(in := 0.0, out1 => "RelatorioUnificado".DosagemAtual[15])
   END_RUNG
   RUNG wire#powerrail
      Contact( "DosagemContinua_DB5".Manual )
   END_RUNG wire#w5
   RUNG wire#powerrail
      Contact( "SinalMisturador2" )
      I_Contact( "DosagemContinua_DB6".Manual )
      Move(in := "SP_Dosagem6", out1 => "RelatorioUnificado".DosagemAtual[16])
   END_RUNG
   RUNG wire#powerrail
      I_Contact( "SinalMisturador2" )
      wire#w6
      Move(in := 0.0, out1 => "RelatorioUnificado".DosagemAtual[16])
   END_RUNG
   RUNG wire#powerrail
      Contact( "DosagemContinua_DB6".Manual )
   END_RUNG wire#w6
   // the same network as SCL:
   "RelatorioUnificado".DosagemAtual[1] := "RegistradorMedidor_DB1".VazaoFiltrada_Lhora;
   "RelatorioUnificado".DosagemAtual[2] := "RegistradorMedidor_DB2".VazaoFiltrada_Lhora;
   "RelatorioUnificado".DosagemAtual[3] := "RegistradorMedidor_DB3".VazaoFiltrada_Lhora;
   "RelatorioUnificado".DosagemAtual[4] := "RegistradorMedidor_DB4".VazaoFiltrada_Lhora;
   "RelatorioUnificado".DosagemAtual[5] := "RegistradorMedidor_DB5".VazaoFiltrada_Lhora;
   "RelatorioUnificado".DosagemAtual[6] := "RegistradorMedidor_DB6".VazaoFiltrada_Lhora;
   IF "SinalTriturador1" AND NOT "DosagemContinua_DB1".Manual THEN
       "RelatorioUnificado".DosagemAtual[11] := "SP_Dosagem1";
   END_IF;
   IF NOT "SinalTriturador1" OR "DosagemContinua_DB1".Manual THEN
       "RelatorioUnificado".DosagemAtual[11] := 0.0;
   END_IF;
   IF "SinalTriturador2" AND NOT "DosagemContinua_DB2".Manual THEN
       "RelatorioUnificado".DosagemAtual[12] := "SP_Dosagem2";
   END_IF;
   IF NOT "SinalTriturador2" OR "DosagemContinua_DB2".Manual THEN
       "RelatorioUnificado".DosagemAtual[12] := 0.0;
   END_IF;
   IF "SinalMisturador1" AND NOT "DosagemContinua_DB3".Manual THEN
       "RelatorioUnificado".DosagemAtual[13] := "SP_Dosagem3";
   END_IF;
   IF NOT "SinalMisturador1" OR "DosagemContinua_DB3".Manual THEN
       "RelatorioUnificado".DosagemAtual[13] := 0.0;
   END_IF;
   IF "SinalMisturador2" AND NOT "DosagemContinua_DB4".Manual THEN
       "RelatorioUnificado".DosagemAtual[14] := "SP_Dosagem4";
   END_IF;
   IF NOT "SinalMisturador2" OR "DosagemContinua_DB4".Manual THEN
       "RelatorioUnificado".DosagemAtual[14] := 0.0;
   END_IF;
   IF "SinalMisturador1" AND NOT "DosagemContinua_DB5".Manual THEN
       "RelatorioUnificado".DosagemAtual[15] := "SP_Dosagem5";
   END_IF;
   IF NOT "SinalMisturador1" OR "DosagemContinua_DB5".Manual THEN
       "RelatorioUnificado".DosagemAtual[15] := 0.0;
   END_IF;
   IF "SinalMisturador2" AND NOT "DosagemContinua_DB6".Manual THEN
       "RelatorioUnificado".DosagemAtual[16] := "SP_Dosagem6";
   END_IF;
   IF NOT "SinalMisturador2" OR "DosagemContinua_DB6".Manual THEN
       "RelatorioUnificado".DosagemAtual[16] := 0.0;
   END_IF;
END_REGION

REGION Network 4: Totalizador Unificado
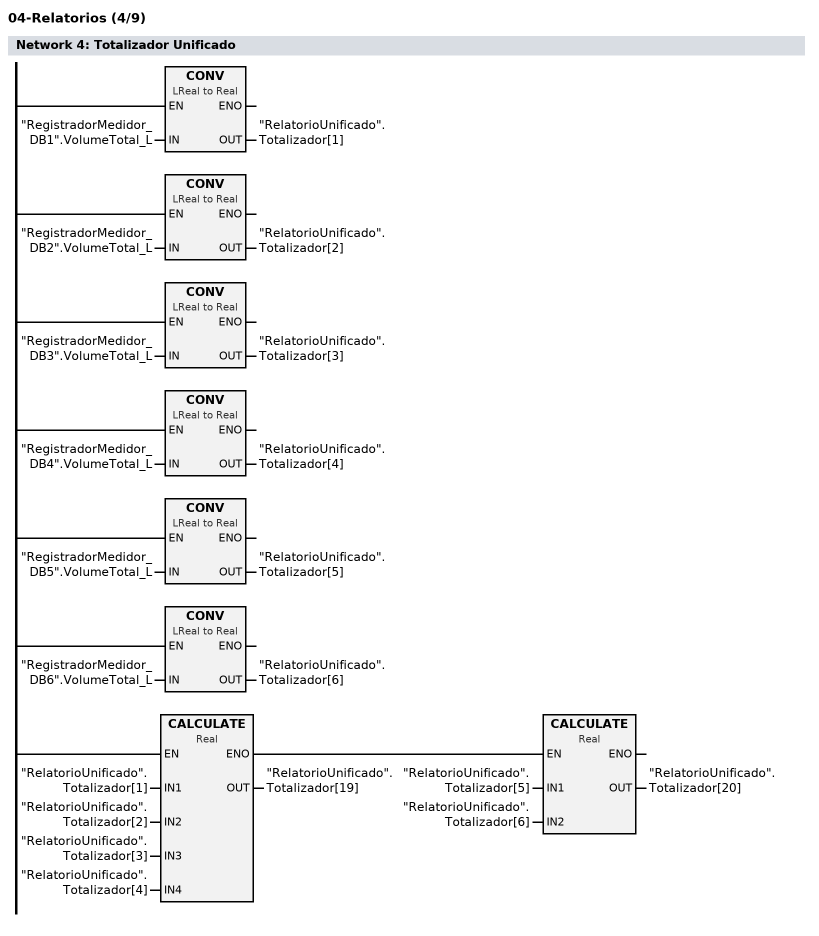
   RUNG wire#powerrail
      { S7_Templates := "[SrcType := LReal, DestType := Real]" } Convert(in := "RegistradorMedidor_DB1".VolumeTotal_L, out => "RelatorioUnificado".Totalizador[1])
   END_RUNG
   RUNG wire#powerrail
      { S7_Templates := "[SrcType := LReal, DestType := Real]" } Convert(in := "RegistradorMedidor_DB2".VolumeTotal_L, out => "RelatorioUnificado".Totalizador[2])
   END_RUNG
   RUNG wire#powerrail
      { S7_Templates := "[SrcType := LReal, DestType := Real]" } Convert(in := "RegistradorMedidor_DB3".VolumeTotal_L, out => "RelatorioUnificado".Totalizador[3])
   END_RUNG
   RUNG wire#powerrail
      { S7_Templates := "[SrcType := LReal, DestType := Real]" } Convert(in := "RegistradorMedidor_DB4".VolumeTotal_L, out => "RelatorioUnificado".Totalizador[4])
   END_RUNG
   RUNG wire#powerrail
      { S7_Templates := "[SrcType := LReal, DestType := Real]" } Convert(in := "RegistradorMedidor_DB5".VolumeTotal_L, out => "RelatorioUnificado".Totalizador[5])
   END_RUNG
   RUNG wire#powerrail
      { S7_Templates := "[SrcType := LReal, DestType := Real]" } Convert(in := "RegistradorMedidor_DB6".VolumeTotal_L, out => "RelatorioUnificado".Totalizador[6])
   END_RUNG
   RUNG wire#powerrail
      { S7_Templates := "SrcType := Real"; S7_Expression := "IN1 + IN2 + IN3 + IN4" } Calculate(in1 := "RelatorioUnificado".Totalizador[1], in2 := "RelatorioUnificado".Totalizador[2], in3 := "RelatorioUnificado".Totalizador[3], in4 := "RelatorioUnificado".Totalizador[4], out => "RelatorioUnificado".Totalizador[19])
      { S7_Templates := "SrcType := Real"; S7_Expression := "IN1 + IN2" } Calculate(in1 := "RelatorioUnificado".Totalizador[5], in2 := "RelatorioUnificado".Totalizador[6], out => "RelatorioUnificado".Totalizador[20])
   END_RUNG
   // the same network as SCL:
   "RelatorioUnificado".Totalizador[1] := LREAL_TO_REAL("RegistradorMedidor_DB1".VolumeTotal_L);
   "RelatorioUnificado".Totalizador[2] := LREAL_TO_REAL("RegistradorMedidor_DB2".VolumeTotal_L);
   "RelatorioUnificado".Totalizador[3] := LREAL_TO_REAL("RegistradorMedidor_DB3".VolumeTotal_L);
   "RelatorioUnificado".Totalizador[4] := LREAL_TO_REAL("RegistradorMedidor_DB4".VolumeTotal_L);
   "RelatorioUnificado".Totalizador[5] := LREAL_TO_REAL("RegistradorMedidor_DB5".VolumeTotal_L);
   "RelatorioUnificado".Totalizador[6] := LREAL_TO_REAL("RegistradorMedidor_DB6".VolumeTotal_L);
   "RelatorioUnificado".Totalizador[19] := "RelatorioUnificado".Totalizador[1] + "RelatorioUnificado".Totalizador[2] + "RelatorioUnificado".Totalizador[3] + "RelatorioUnificado".Totalizador[4];
   "RelatorioUnificado".Totalizador[20] := "RelatorioUnificado".Totalizador[5] + "RelatorioUnificado".Totalizador[6];
END_REGION

